(* 상대 PLC 끊김 / 통신 한쪽 고장 *)
_fbRedPeerLost(i_stEntry := TC_EVENTS.PmsSystem.RedPeerLost, i_bActive := i_bRedUse AND i_ePeer = E_RedPeer.Lost, i_nArgs := 0, i_asArg := _asArg);
IF _fbRedLinkFault.q_bRaised <> (i_bRedUse AND (i_ePeer = E_RedPeer.EapLost OR i_ePeer = E_RedPeer.WireLost)) THEN
	IF i_ePeer = E_RedPeer.EapLost THEN
		_asArg[1] := "EAP";
	ELSE
		_asArg[1] := "접점";
	END_IF
END_IF
_fbRedLinkFault(i_stEntry := TC_EVENTS.PmsSystem.RedLinkFault, i_bActive := i_bRedUse AND (i_ePeer = E_RedPeer.EapLost OR i_ePeer = E_RedPeer.WireLost), i_nArgs := 1, i_asArg := _asArg);

(* 동기화 값을 못 받음: EAP는 살아 있는데 동기화 값이 5 s 넘게 안 옴 *)
_tonRedSync(IN := i_bRedUse AND i_bPeerEapOk AND NOT i_bSyncFresh, PT := T#5S);
_fbRedSyncLost(i_stEntry := TC_EVENTS.PmsSystem.RedSyncLost, i_bActive := _tonRedSync.Q, i_nArgs := 0, i_asArg := _asArg);

(* 이중화 설정 오류: 두 PLC 역할이 같거나 Net ID가 RED_SET과 안 맞음 *)
IF _fbRedFailed.q_bRaised <> (i_eRedState = E_RedState.Failed) THEN
	IF i_bRoleConflict THEN
		_asArg[1] := "두 PLC의 역할이 같음";
	ELSE
		_asArg[1] := "이 PLC의 Net ID가 RED_SET과 맞지 않음";
	END_IF
END_IF
_fbRedFailed(i_stEntry := TC_EVENTS.PmsSystem.RedFailed, i_bActive := i_eRedState = E_RedState.Failed, i_nArgs := 1, i_asArg := _asArg);

(* 동기화로 설정을 맞춤 (Active가 바꾼 설정이 이 PLC에 반영됨) *)
IF i_nSyncApplied <> _nRedAppliedLast THEN
	_asArg[1] := TO_WSTRING(i_nSyncApplied - _nRedAppliedLast);
	_nRedAppliedLast := i_nSyncApplied;
	_fbRedSyncApplied.M_SendEvent(1, _asArg);
END_IF
END_ACTION

ACTION A_LogProtection:
// 보호 알람
(* ===== 1) 보호 (알람: 발생·해소 1회씩). 규칙 칸·대상마다. 심각도는 처음 만들 때 조치 기준 ===== *)
FOR _i := 1 TO GVL_PARAM.RULE_COUNT DO
	_m := 0;
	IF iq_aipRule[_i] <> 0 THEN _m := iq_aipRule[_i].ModuleId; END_IF
	FOR _t := 1 TO GVL_PARAM.PROT_TARGET_MAX DO
		// [결함 8 수정 2026-11-03: 대응 칸이 비면 조치가 안 걸리므로 문구·심각도도 조치 없음 (알람만). 원래는 설정 stProt를 그대로 씀:
		//   M_FillProtArgs(..., iq_astRuleCfg[_i].stProt, _asArg) / M_ProtEventBySeverity(iq_astRuleCfg[_i].stProt)]
		_stProtTxt := iq_astRuleCfg[_i].stProt;
		IF iq_aipResp[_i] = 0 THEN
			_stProtTxt.ePcsAction	:= E_PcsAction.None;
			_stProtTxt.eBatAction	:= E_BatAction.None;
			_stProtTxt.eModeAction	:= E_ModeAction.None;
			_stProtTxt.fPPct		:= 100.0;
			_stProtTxt.fQPct		:= 100.0;
		END_IF
		IF _aafbRule[_i, _t].q_bRaised <> iq_aabRule[_i, _t] THEN
			M_FillProtArgs(_m, M_RuleTarget(iq_astRuleCfg[_i].eScope, _t), _stProtTxt, _asArg);
		END_IF
		_aafbRule[_i, _t](i_stEntry := M_ProtEventBySeverity(_stProtTxt), i_bActive := iq_aabRule[_i, _t], i_nArgs := 5, i_asArg := _asArg);
	END_FOR
END_FOR

(* ===== BMS 명령 실패 (알람, 잠그지 않음). 이벤트 항목은 PmsProt.BatLocked를 씀 (문구는 이벤트 클래스에서) ===== *)
FOR _m := 1 TO GVL_PARAM.BMS_COUNT DO
	IF _afbBmsCmdFail[_m].q_bRaised <> (iq_aeBmsFailCmd[_m] <> E_BatCmd.None) THEN
		_asArg[1] := TO_WSTRING(_m);
		_asArg[2] := WCONCAT(F_TxtBatCmd(iq_aeBmsFailCmd[_m]), " 명령 접수 안 됨");
	END_IF
	_afbBmsCmdFail[_m](i_stEntry := TC_EVENTS.PmsProt.BatLocked, i_bActive := iq_aeBmsFailCmd[_m] <> E_BatCmd.None, i_nArgs := 2, i_asArg := _asArg);
END_FOR

(* ===== 가상신호 (알람): 종류가 바뀌면(전압 → 유효전력 등) 해소 후 새 종류로 다시 발생 ===== *)
FOR _g := 1 TO GVL_PARAM.GROUP_COUNT DO
	_nVirtualKind := SEL(i_bTestMode AND iq_astVirtual[_g].bVEna, 0, 1) + SEL(i_bTestMode AND iq_astVirtual[_g].bPEna, 0, 2);
	IF _nVirtualKind <> _anVirtualKind[_g] THEN
		IF _afbVirtual[_g].q_bRaised THEN
			_afbVirtual[_g](i_stEntry := TC_EVENTS.PmsOutput.VirtualOn, i_bActive := FALSE, i_nArgs := 0, i_asArg := _asArg);
		END_IF
		_asArg[1] := TO_WSTRING(_g);
		CASE _nVirtualKind OF
			1:	_asArg[2] := "전압";
			2:	_asArg[2] := "유효전력";
			3:	_asArg[2] := "전압·유효전력";
		END_CASE
		_anVirtualKind[_g] := _nVirtualKind;
	END_IF
	_afbVirtual[_g](i_stEntry := TC_EVENTS.PmsOutput.VirtualOn, i_bActive := _nVirtualKind <> 0, i_nArgs := 2, i_asArg := _asArg);
END_FOR

// 보호가 요청 모드를 Manual로 바꿈 (메시지, 보호가 걸릴 때마다 1회. 걸려 있는 동안 Auto 재요청을 되돌려도 다시 남기지 않음)
FOR _u := 1 TO GVL_PARAM.UNIT_COUNT DO
	IF iq_abModeForced[_u] AND NOT _abModeForcedLogged[_u] THEN
		_asArg[1] := TO_WSTRING(_u);
		_asArg[2] := M_ModuleName(iq_astUnitProt[_u].nModeModule);
		_asArg[3] := TO_WSTRING(iq_astUnitProt[_u].nModeModule);
		_fbModeForced.M_SendEvent(3, _asArg);
		_abModeForcedLogged[_u] := TRUE;
	END_IF
	IF NOT iq_astUnitProt[_u].bModeManualReq THEN
		_abModeForcedLogged[_u] := FALSE;
	END_IF
END_FOR
END_ACTION

ACTION A_LogDeviceFail:
// 명령 실패·장비 쓰기 실패
(* ===== 2) 명령 실패 (알람) ===== *)
FOR _u := 1 TO GVL_PARAM.UNIT_COUNT DO
	IF _afbCmdFail[_u].q_bRaised <> (iq_aeFailCmd[_u] <> E_PcsCmd.None) THEN
		_asArg[1] := TO_WSTRING(_u);
		_asArg[2] := F_TxtPcsCmd(iq_aeFailCmd[_u]);
	END_IF
	_afbCmdFail[_u](i_stEntry := TC_EVENTS.PmsSeq.CmdFail, i_bActive := iq_aeFailCmd[_u] <> E_PcsCmd.None, i_nArgs := 2, i_asArg := _asArg);
END_FOR

(* ===== 2-0) 장비 쓰기 실패 (알람): 드라이버가 상태 bWriteFail로 알림 (FB_DeviceBase.M_MarkWriteResult) ===== *)
FOR _u := 1 TO GVL_PARAM.UNIT_COUNT DO
	IF _afbUnitWriteFail[_u].q_bRaised <> iq_astUnit[_u].bWriteFail THEN
		_asArg[1] := F_TxtNum("유닛 ", _u);
	END_IF
	_afbUnitWriteFail[_u](i_stEntry := TC_EVENTS.PmsSystem.WriteFail, i_bActive := iq_astUnit[_u].bWriteFail, i_nArgs := 1, i_asArg := _asArg);
END_FOR
FOR _m := 1 TO GVL_PARAM.BMS_COUNT DO
	IF _afbBmsWriteFail[_m].q_bRaised <> iq_astBms[_m].bWriteFail THEN
		_asArg[1] := F_TxtNum("BMS ", _m);
	END_IF
	_afbBmsWriteFail[_m](i_stEntry := TC_EVENTS.PmsSystem.WriteFail, i_bActive := iq_astBms[_m].bWriteFail, i_nArgs := 1, i_asArg := _asArg);
END_FOR
END_ACTION

ACTION A_LogSource:
// 지령원 요청·끊김, 코어 상태 요청
(* ===== 3) 지령원: 상태 변경 요청(메시지), 끊김(알람) ===== *)
FOR _i := 1 TO GVL_PARAM.SOURCE_COUNT DO
	IF iq_aipSource[_i] <> 0 AND_THEN iq_astSrcOut[_i].bValid THEN
		_asArg[1] := STRING_TO_WSTRING(iq_aipSource[_i].ModuleName);
		_asArg[2] := TO_WSTRING(iq_aipSource[_i].ModuleId);
		// PCS 요청: 받은 것은 지금 요청과 다를 때만(Reset은 항상), 운전 모드 설정 때문에 무시한 것은 지령 무시로
		IF iq_astSrcOut[_i].stPcsReq.eCmd <> E_PcsCmd.None THEN
			_asArg[3] := F_TxtPcsCmd(iq_astSrcOut[_i].stPcsReq.eCmd);
			IF iq_astSrcOut[_i].stPcsReq.nUnit = 0 THEN
				_asArg[4] := "전체";
			ELSE
				_asArg[4] := F_TxtNum("유닛 ", iq_astSrcOut[_i].stPcsReq.nUnit);
			END_IF
			IF iq_abPcsReqTaken[_i] OR iq_astSrcOut[_i].stPcsReq.eCmd = E_PcsCmd.Reset THEN
				IF iq_astSrcOut[_i].stPcsReq.eCmd <> _aeLastPcsReq[_i] OR iq_astSrcOut[_i].stPcsReq.nUnit <> _anLastPcsUnit[_i]
					OR iq_astSrcOut[_i].stPcsReq.eCmd = E_PcsCmd.Reset THEN
					_fbStateReq.M_SendEvent(4, _asArg);
					_aeLastPcsReq[_i]	:= iq_astSrcOut[_i].stPcsReq.eCmd;
					_anLastPcsUnit[_i]	:= iq_astSrcOut[_i].stPcsReq.nUnit;
				END_IF
			ELSIF i_stSet.bCmdRefused THEN
				_asArg[3] := WCONCAT(_asArg[3], WCONCAT(" ", _asArg[4]));
				_asArg[4] := "이 운전 모드에서 받지 않음 (stStateMode·모드 전환)";
				_fbCmdRefused.M_SendEvent(4, _asArg);
			END_IF
		END_IF
		// 배터리 요청: 받은 것은 항상, 무시한 것은 지령 무시로. Reset은 운전 모드와 관계없이 시퀀서가 보내므로 받은 것으로 기록 (PCS Reset과 같음)
		IF iq_astSrcOut[_i].stBatReq.eCmd <> E_BatCmd.None THEN
			_asArg[3] := F_TxtBatCmd(iq_astSrcOut[_i].stBatReq.eCmd);
			IF iq_astSrcOut[_i].stBatReq.nBatGroup = 0 THEN
				_asArg[4] := "전체";
			ELSE
				_asArg[4] := F_TxtNum("배터리 그룹 ", iq_astSrcOut[_i].stBatReq.nBatGroup);
			END_IF
			IF iq_abBatReqTaken[_i] OR iq_astSrcOut[_i].stBatReq.eCmd = E_BatCmd.Reset THEN
				_fbStateReq.M_SendEvent(4, _asArg);
			ELSIF i_stSet.bCmdRefused THEN
				_asArg[3] := WCONCAT(_asArg[3], WCONCAT(" ", _asArg[4]));
				_asArg[4] := "이 운전 모드에서 받지 않음 (stStateMode)";
				_fbCmdRefused.M_SendEvent(4, _asArg);
			END_IF
		END_IF
	END_IF

	IF iq_astSrcOut[_i].bValid THEN
		_abEverValid[_i] := TRUE;
	END_IF
	// [9번 수정 2026-11-09: 등록 bLostAlarm FALSE면 알람 안 냄 (EMS → 브로커 끊김 알람으로 대신). 원래 조건에 bLostAlarm 없음]
	_bLost := iq_aipSource[_i] <> 0 AND_THEN (iq_astReg[_i].bEnable AND iq_astReg[_i].bLostAlarm AND _abEverValid[_i] AND NOT iq_astSrcOut[_i].bValid);
	IF _afbSrcLost[_i].q_bRaised <> _bLost AND iq_aipSource[_i] <> 0 THEN
		_asArg[1] := STRING_TO_WSTRING(iq_aipSource[_i].ModuleName);
		_asArg[2] := TO_WSTRING(iq_aipSource[_i].ModuleId);
	END_IF
	_afbSrcLost[_i](i_stEntry := TC_EVENTS.PmsOutput.SourceLost, i_bActive := _bLost, i_nArgs := 2, i_asArg := _asArg);
END_FOR
END_ACTION

ACTION A_LogRefused:
// 무시한 지령·기동 조건 대기·지령값 이상·배터리 요청 거부
(* ===== 3-2) 무시한 지령 (메시지): 이상값(지령원별), 방향 반대(유닛별). 새로 생길 때 1회 ===== *)
FOR _i := 1 TO GVL_PARAM.SOURCE_COUNT DO
	IF i_stSet.bCmdRefused AND iq_abBadValue[_i] AND NOT _abLastBad[_i] AND iq_aipSource[_i] <> 0 THEN
		_asArg[1] := STRING_TO_WSTRING(iq_aipSource[_i].ModuleName);
		_asArg[2] := TO_WSTRING(iq_aipSource[_i].ModuleId);
		_asArg[3] := "지령값";
		// [결함 9 수정 2026-11-03: NaN을 비교하지 않고 비트로 봄 (원래 IF iq_afBadValue[_i] <> iq_afBadValue[_i] THEN → FPU 예외)]
		MEMCPY(ADR(_dwBadBits), ADR(iq_afBadValue[_i]), SIZEOF(_dwBadBits));
		IF (_dwBadBits AND 16#7F800000) = 16#7F800000 AND (_dwBadBits AND 16#007FFFFF) <> 0 THEN
			_asArg[4] := "이상값 (숫자 아님)";
		ELSIF (_dwBadBits AND 16#7F800000) = 16#7F800000 OR_ELSE ABS(iq_afBadValue[_i]) >= 1.0E9 THEN
			_asArg[4] := "이상값 (너무 큼)";
		ELSE
			_asArg[4] := WCONCAT("이상값 ", TO_WSTRING(F_RealToDint(iq_afBadValue[_i])));	// [결함 13 수정 2026-11-04: REAL_TO_DINT → F_RealToDint]
		END_IF
		_fbCmdRefused.M_SendEvent(4, _asArg);
	END_IF
	_abLastBad[_i] := iq_abBadValue[_i];
END_FOR
FOR _u := 1 TO GVL_PARAM.UNIT_COUNT DO
	IF i_stSet.bCmdRefused AND iq_aeManualRefuse[_u] <> _aeLastCmdRefuse[_u] AND iq_aeManualRefuse[_u] = E_CmdRefuse.Reversed THEN
		_asArg[1] := M_ModuleName(iq_anManualRefuseModule[_u]);
		_asArg[2] := TO_WSTRING(iq_anManualRefuseModule[_u]);
		_asArg[3] := F_TxtNum("유닛 ", _u);
		_asArg[4] := "방향 반대 (운전 중인 방향과 다름, 앞 값 유지)";
		_fbCmdRefused.M_SendEvent(4, _asArg);
	END_IF
	_aeLastCmdRefuse[_u] := iq_aeManualRefuse[_u];
END_FOR

(* ===== 3-2-1) 기동 조건 대기 (메시지): 대기가 시작되거나 막은 모듈·이유가 바뀔 때 1회 ===== *)
FOR _g := 1 TO GVL_PARAM.GROUP_COUNT DO
	IF iq_abWaitPermit[_g] AND NOT iq_abPermit[_g] THEN
		IF NOT _abPermitLogged[_g] OR iq_anPermitModule[_g] <> _anPermitModule[_g] OR iq_anPermitReason[_g] <> _anPermitReason[_g] THEN
			_asArg[1] := TO_WSTRING(_g);
			_asArg[2] := M_ModuleName(iq_anPermitModule[_g]);
			_asArg[3] := M_ReasonText(iq_anPermitModule[_g], iq_anPermitReason[_g]);
			_asArg[4] := TO_WSTRING(iq_anPermitModule[_g]);
			_fbPermitWait.M_SendEvent(4, _asArg);
			_abPermitLogged[_g]	:= TRUE;
			_anPermitModule[_g]	:= iq_anPermitModule[_g];
			_anPermitReason[_g]	:= iq_anPermitReason[_g];
		END_IF
	ELSE
		_abPermitLogged[_g] := FALSE;
	END_IF
END_FOR

(* ===== 3-2-2) 지령값 이상 (메시지): 디스패처가 NaN·무한대를 0으로 바꾼 유닛, 생길 때 1회 ===== *)
FOR _u := 1 TO GVL_PARAM.UNIT_COUNT DO
	IF iq_abBadSet[_u] AND NOT _abLastBadSet[_u] THEN
		_asArg[1] := TO_WSTRING(_u);
		_fbBadSet.M_SendEvent(1, _asArg);
	END_IF
	_abLastBadSet[_u] := iq_abBadSet[_u];
END_FOR

(* ===== 3-3) 배터리 요청 거부 (메시지): 거부된 요청마다 1회 ===== *)
FOR _b := 1 TO GVL_PARAM.BAT_COUNT DO
	IF i_stSet.bBatRefused AND iq_abBatRefusedNow[_b] THEN
		_asArg[1] := F_TxtNum("배터리 그룹 ", _b);
		IF iq_aeBatRefuse[_b] = E_SeqRefuse.UnitRunning THEN
			_asArg[2] := "배터리 개방";
			_asArg[3] := "버스의 유닛이 운전 중 (정지 후 개방)";
		ELSE
			_asArg[2] := "배터리";
			_asArg[3] := F_TxtRefuse(iq_aeBatRefuse[_b]);
		END_IF
		_fbRefused.M_SendEvent(3, _asArg);
	END_IF
END_FOR
END_ACTION

ACTION A_LogOutput:
// 출력 제한, 자세한 기록
(* ===== 4) 출력 제한: 이유(단계·모듈·이유)가 바뀌고 유지 시간이 지나야 기록 ===== *)
FOR _g := 1 TO GVL_PARAM.GROUP_COUNT DO
	IF NOT M_SameLimitReason(iq_astAutoPDiag[_g], _astCand[_g]) THEN
		_astCand[_g] := iq_astAutoPDiag[_g];
		_atonHold[_g](IN := FALSE);
	END_IF
	_atonHold[_g](IN := NOT M_SameLimitReason(_astCand[_g], _astLogged[_g]), PT := i_stSet.tHold);
	IF _atonHold[_g].Q THEN
		IF M_IsLoggedStage(_astCand[_g].eStage) THEN
			_asArg[1] := TO_WSTRING(_g);
			_asArg[2] := F_TxtStage(_astCand[_g].eStage);
			IF _astCand[_g].eStage = E_DiagStage.UnitLimit THEN
				_asArg[3] := F_TxtLimitBy(_astCand[_g].eUnitBy);
			ELSE
				_asArg[3] := M_ReasonText(_astCand[_g].nModule, _astCand[_g].nReason);
			END_IF
			_asArg[4] := TO_WSTRING(_astCand[_g].nModule);
			_asArg[5] := TO_WSTRING(F_RealToDint(iq_astAutoPDiag[_g].fReq));	// [결함 13 수정 2026-11-04: REAL_TO_DINT → F_RealToDint (NaN·범위 밖 예외 없음)]
			_asArg[6] := TO_WSTRING(F_RealToDint(iq_astAutoPDiag[_g].fOut));
			_fbLimited.M_SendEvent(6, _asArg);
		ELSIF M_IsLoggedStage(_astLogged[_g].eStage) THEN
			_asArg[1] := TO_WSTRING(_g);
			_fbFree.M_SendEvent(1, _asArg);
		END_IF
		_astLogged[_g] := _astCand[_g];
		_atonHold[_g](IN := FALSE);
	END_IF
END_FOR

(* ===== 5) 자세한 기록 (설정으로 켬) ===== *)
FOR _u := 1 TO GVL_PARAM.UNIT_COUNT DO
	IF i_stSet.bUnitLimited AND iq_astUnitDiag[_u].ePBy <> _aeLastLimBy[_u]
		AND iq_astUnitDiag[_u].ePBy <> E_UnitLimitBy.NotRun AND iq_astUnitDiag[_u].ePBy <> E_UnitLimitBy.NotAvail THEN
		_asArg[1] := TO_WSTRING(_u);
		_asArg[2] := F_TxtLimitBy(iq_astUnitDiag[_u].ePBy);
		_asArg[3] := TO_WSTRING(F_RealToDint(iq_astUnitDiag[_u].fPReq));	// [결함 13 수정 2026-11-04: REAL_TO_DINT → F_RealToDint]
		_asArg[4] := TO_WSTRING(F_RealToDint(iq_astUnitDiag[_u].fPOut));
		_fbUnitLim.M_SendEvent(4, _asArg);
	END_IF
	_aeLastLimBy[_u] := iq_astUnitDiag[_u].ePBy;

	IF i_stSet.bReqRefused AND iq_aeRefuse[_u] <> _aeLastRefuse[_u] AND iq_aeRefuse[_u] <> E_SeqRefuse.None THEN
		_asArg[1] := F_TxtNum("유닛 ", _u);
		_asArg[2] := "기동";
		_asArg[3] := F_TxtRefuse(iq_aeRefuse[_u]);
		_fbRefused.M_SendEvent(3, _asArg);
	END_IF
	_aeLastRefuse[_u] := iq_aeRefuse[_u];

	IF i_stSet.bSeqChange AND iq_aeUnitSeq[_u] <> _aeLastSeq[_u] THEN
		_asArg[1] := TO_WSTRING(_u);
		_asArg[2] := F_TxtSeq(_aeLastSeq[_u]);
		_asArg[3] := F_TxtSeq(iq_aeUnitSeq[_u]);
		_fbSeqChange.M_SendEvent(3, _asArg);
	END_IF
	_aeLastSeq[_u] := iq_aeUnitSeq[_u];

	IF i_stSet.bModeChange AND iq_aeOpMode[_u] <> _aeLastMode[_u] THEN
		_asArg[1] := TO_WSTRING(_u);
		_asArg[2] := F_TxtOpMode(_aeLastMode[_u]);
		_asArg[3] := F_TxtOpMode(iq_aeOpMode[_u]);
		_fbModeChange.M_SendEvent(3, _asArg);
	END_IF
	_aeLastMode[_u] := iq_aeOpMode[_u];
END_FOR
END_ACTION

END_FUNCTION_BLOCK

// ---- 10_Core/30_Request/FB_CtrlModeMgr.TcPOU
FUNCTION_BLOCK FB_CtrlModeMgr EXTENDS FB_SourceBase		// 제어 모드 관리자: 등록한 제어 모드(I_ControlMode) 중 하나만 켜고 전환을 맡음. 코어에는 지령원 하나로 보임
// 등록: GVL_SITE.g_aipSource 한 칸 + GVL_PERSIST.g_astSourceReg 같은 칸 (ePowerMode := Auto → Auto 유닛에만 적용). 상태 요청(Run·Stop 등)·제한은 내지 않음
// 요청(i_nModeReq = 모드 칸 번호, 0 = 모드 없음)이 바뀌면: 진입 검사 → 지금 모드 M_Exit → (출력 0 → 지연) → 진입 검사 다시 → 새 모드 M_Enter. 시작한 전환은 끝까지 진행
// 진입 검사에 걸리면 지금 모드를 그대로 둠. 켜진 모드가 스스로 끝내면(bExitReq) 대체 모드(i_stSet.nFallback)로
// 처리한 요청값은 다시 처리하지 않음 (거부·스스로 끝남 뒤 저절로 다시 들어가지 않게). 같은 값을 다시 시도하려면 i_bRetry
// 단위: i_nUnit = 0 → 그룹 하나를 맡음 (그룹 지령 fPSet, 모드는 그룹 값을 봄. 그룹이 2개 이상이면 그룹마다 인스턴스, 등록표 nGroup)
//       i_nUnit = n → 유닛(PCS) n만 맡음 (유닛별 값 astUnit[n], 모드는 FB_UnitView 유닛 값을 봄). PCS마다 관리자 하나 + 모드 인스턴스 한 세트 + 설정 한 세트
//       유닛 단위의 접속점 값은 i_stSet.ePccShare (같은 접속점을 여러 유닛이 쓰면 몫으로 나눔). 접속점이 따로면 유닛마다 제어 그룹을 따로 둠 (GVL_SITE.GROUP_CFG)
// 모드는 FB_ModuleList에 없으므로 설정 점검(M_CheckSet)은 이 FB가 대신 부름
VAR_INPUT
	i_aipMode	: ARRAY[1..GVL_PARAM.CTRL_MODE_COUNT] OF I_ControlMode;	// 등록한 제어 모드 (MAIN 액션 A_PassModuleSet이 GVL_SITE.g_aipCtrlModeN을 매 스캔 넘김). 빈 칸 = 0
	i_stSet		: ST_CtrlModeSet;	// 전환 설정 (A_PassModuleSet이 GVL_PERSIST.g_stModuleSet 칸을 매 스캔 넘김)
	i_nModeReq	: UINT;				// 요청 모드 칸 번호. 0 = 모드 없음 (지령을 내지 않음)
	i_bRetry	: BOOL;				// 같은 요청값을 다시 처리 (쓰면 한 번 처리하고 FALSE로 돌아감)
	i_stTime	: ST_LocalTime;		// 현지 시각 (MAIN 액션 A_PassModuleSet이 매 스캔 넘김). 시간표를 쓰는 모드가 봄
	i_nUnit		: UINT;				// 0 = 그룹 단위. 1~ = 이 유닛(PCS) 단위. 선언에서 정함 (GVL_SITE)
	i_pUnitView	: POINTER TO ARRAY[1..GVL_PARAM.UNIT_COUNT] OF ST_UnitView;	// 유닛 단위일 때: MAIN.fbUnitView.q_astView 주소 (A_PassModuleSet이 매 스캔 넘김). 0 = 연결 안 됨
END_VAR
VAR_OUTPUT
	q_nActive		: UINT;					// 켜진 모드 칸 번호. 0 = 없음 (전환 중에도 0)
	q_sActive		: STRING(31);			// 켜진 모드 이름 (ModuleName)
	q_eStep			: E_CtrlModeStep;		// 관리자 단계
	q_nTarget		: UINT;					// 전환 중 목표 칸 번호 (Leaving일 때만, 0 = 모드 없음으로 가는 중)
	q_eRefuse		: E_CtrlModeRefuse;		// 마지막으로 처리한 요청의 결과 (None = 접수)
	q_nRefuseReason	: UINT;					// NotReady일 때 그 모드의 이유 코드 (M_ModeReasonText)
	q_nExitSlot		: UINT;					// 마지막으로 스스로 끝낸 모드 칸 번호
	q_nExitReason	: UINT;					// 그 이유 코드 (M_ModeReasonText)
	q_bChanged		: BOOL;					// 켜진 모드가 바뀐 스캔 (1스캔, 기록용)
	q_bRefusedNow	: BOOL;					// 이번 스캔에 요청을 거부함 (1스캔, 기록용). 칸 q_nRefuseSlot, 결과 q_eRefuse·q_nRefuseReason [7번 수정 2026-11-09: 추가]
	q_nRefuseSlot	: UINT;					// 마지막으로 거부한 요청 칸 번호
	q_bExitedNow	: BOOL;					// 이번 스캔에 켜진 모드가 스스로 끝남 (1스캔, 기록용). 칸 q_nExitSlot, 이유 q_nExitReason [7번 수정 2026-11-09: 추가]
	q_fPccP			: REAL;					// kW, 모드가 본 접속점 P (공급 +). 유닛 단위면 ePccShare를 적용한 값
END_VAR
VAR
	_nHandledReq	: UINT;				// 처리를 끝낸 요청값 (요청이 이것과 다를 때만 새로 처리)
	_nActive		: UINT;				// 켜진 모드 칸 번호
	_nTarget		: UINT;				// 진행 중인 전환의 목표 (끝날 때까지 고정)
	_bLeaveP		: BOOL;				// 전환 중 P를 0으로 냄 (이전 모드가 P를 내던 경우만)
	_bLeaveQ		: BOOL;				// 전환 중 Q를 0으로 냄
	_bPrevP			: BOOL;				// 켜진 모드가 지난 스캔에 P를 냄
	_bPrevQ			: BOOL;
	_tonZero		: TON;
	_stModeOut		: ST_CtrlModeOut;	// 켜진 모드의 이번 스캔 결과
	_stModeView		: ST_CtrlModeView;	// 모드에 넘기는 값 (이번 스캔)
	(* [16번 수정 2026-11-09: 추가] 유닛별 값을 내는 모드(bUnitOut)의 전환 중 0 *)
	_bPrevUnitOut	: BOOL;				// 켜진 모드가 지난 스캔에 유닛별 값을 냄
	_abPrevUnitP	: ARRAY[1..GVL_PARAM.UNIT_COUNT] OF BOOL;
	_abPrevUnitQ	: ARRAY[1..GVL_PARAM.UNIT_COUNT] OF BOOL;
	_bLeaveUnit		: BOOL;				// 전환 중 유닛 칸으로 0을 냄 (이전 모드가 유닛별 값을 내던 경우)
	_abLeaveUnitP	: ARRAY[1..GVL_PARAM.UNIT_COUNT] OF BOOL;
	_abLeaveUnitQ	: ARRAY[1..GVL_PARAM.UNIT_COUNT] OF BOOL;
END_VAR

METHOD M_UpdateOutput : BOOL
VAR
	stNoMode	: ST_CtrlModeOut;
	stOld		: ST_SourceOutput;	// 지난 스캔 낸 값 (새 지령 판단)
	bNew		: BOOL;
	stNoReq		: ST_UnitReq;
	k			: UINT;
	nCode		: UINT;
	nFallback	: UINT;
	bOk			: BOOL;
END_VAR
q_bChanged	:= FALSE;
q_bRefusedNow	:= FALSE;
q_bExitedNow	:= FALSE;
IF i_nUnit = 0 THEN
	_stModeView.stGroup	:= _stView;		// FB_SourceBase가 이번 스캔 채운 대상 그룹 값
ELSE
	_stModeView.stGroup	:= M_UnitView();	// 이 유닛 값 (접속점은 ePccShare 몫)
END_IF
_stModeView.stTime	:= i_stTime;
q_fPccP := _stModeView.stGroup.stPcc.stMeas.stP.fValue;

// 0) 켜진 모드가 등록에서 빠졌으면 (온라인 변경) 모드 없음으로
IF q_eStep = E_CtrlModeStep.Active AND NOT M_Valid(i_nSlot := _nActive) THEN
	_nActive	:= 0;
	q_eStep		:= E_CtrlModeStep.Idle;
	q_bChanged	:= TRUE;
END_IF

// 1) 새 요청 (전환 중이면 끝난 뒤 처리)
IF q_eStep <> E_CtrlModeStep.Leaving AND (i_nModeReq <> _nHandledReq OR i_bRetry) THEN
	_nHandledReq	:= i_nModeReq;
	q_eRefuse		:= E_CtrlModeRefuse.None;
	q_nRefuseReason	:= 0;
	IF i_nModeReq <> _nActive THEN
		IF i_nModeReq <> 0 AND NOT M_Valid(i_nSlot := i_nModeReq) THEN
			q_eRefuse := E_CtrlModeRefuse.BadSlot;
			q_nRefuseSlot	:= i_nModeReq;
			q_bRefusedNow	:= TRUE;
		ELSE
			nCode := 0;
			IF i_nModeReq <> 0 THEN
				nCode := i_aipMode[i_nModeReq].M_CheckEnter(i_stView := _stModeView);
			END_IF
			IF nCode = 0 THEN
				M_StartSwitch(i_nTarget := i_nModeReq);
			ELSE
				q_eRefuse		:= E_CtrlModeRefuse.NotReady;	// 지금 모드는 그대로
				q_nRefuseReason	:= nCode;
				q_nRefuseSlot	:= i_nModeReq;
				q_bRefusedNow	:= TRUE;
			END_IF
		END_IF
	END_IF
	i_bRetry := FALSE;		// 처리한 뒤에만 지움 (전환 중에 온 재시도는 끝난 뒤 처리)
END_IF

// 2) 전환 중: 0으로 둔 시간이 지나면 진입 검사를 다시 하고 새 모드로 (지연 동안 조건이 바뀌었을 수 있음)
_tonZero(IN := q_eStep = E_CtrlModeStep.Leaving, PT := i_stSet.tZeroDelay);
IF q_eStep = E_CtrlModeStep.Leaving AND _tonZero.Q THEN
	bOk := TRUE;
	IF _nTarget <> 0 THEN
		IF M_Valid(i_nSlot := _nTarget) THEN
			nCode := i_aipMode[_nTarget].M_CheckEnter(i_stView := _stModeView);
			IF nCode <> 0 THEN
				bOk				:= FALSE;
				q_eRefuse		:= E_CtrlModeRefuse.NotReady;
				q_nRefuseReason	:= nCode;
			END_IF
		ELSE
			bOk				:= FALSE;
			q_eRefuse		:= E_CtrlModeRefuse.BadSlot;
			q_nRefuseReason	:= 0;
		END_IF
		IF NOT bOk THEN
			q_nRefuseSlot	:= _nTarget;
			q_bRefusedNow	:= TRUE;
		END_IF
	END_IF
	IF bOk THEN
		M_EnterMode(i_nSlot := _nTarget);
	ELSE
		M_EnterMode(i_nSlot := 0);
	END_IF
END_IF

// 3) 켜진 모드 계산. 스스로 끝내면 대체 모드로
IF q_eStep = E_CtrlModeStep.Active THEN
	_bPrevP		:= _stModeOut.bPSetActive;		// 지난 스캔에 내던 쪽 (끝내는 스캔에 지령을 비워도 0으로 둘 수 있게)
	_bPrevQ		:= _stModeOut.bQSetActive;
	_bPrevUnitOut	:= _stModeOut.bUnitOut;
	FOR k := 1 TO GVL_PARAM.UNIT_COUNT DO
		_abPrevUnitP[k]	:= _stModeOut.bUnitOut AND _stModeOut.astUnit[k].bPSetActive;
		_abPrevUnitQ[k]	:= _stModeOut.bUnitOut AND _stModeOut.astUnit[k].bQSetActive;
	END_FOR
	_stModeOut	:= i_aipMode[_nActive].M_Calc(i_stView := _stModeView);
	IF _stModeOut.bExitReq THEN
		q_nExitSlot		:= _nActive;
		q_nExitReason	:= _stModeOut.nReason;
		q_bExitedNow	:= TRUE;
		nFallback		:= 0;
		IF i_stSet.nFallback <> _nActive AND M_Valid(i_nSlot := i_stSet.nFallback) THEN
			IF i_aipMode[i_stSet.nFallback].M_CheckEnter(i_stView := _stModeView) = 0 THEN
				nFallback := i_stSet.nFallback;
			END_IF
		END_IF
		M_StartSwitch(i_nTarget := nFallback);
		// 대체 모드로 바로 들어갔으면 이번 스캔 값을 냄 (그 모드의 bExitReq는 다음 스캔에 봄)
		IF q_eStep = E_CtrlModeStep.Active THEN
			_stModeOut := i_aipMode[_nActive].M_Calc(i_stView := _stModeView);
		END_IF
	END_IF
ELSIF q_eStep = E_CtrlModeStep.Idle THEN
	_stModeOut	:= stNoMode;
	_bPrevP		:= FALSE;
	_bPrevQ		:= FALSE;
	_bPrevUnitOut	:= FALSE;
	FOR k := 1 TO GVL_PARAM.UNIT_COUNT DO
		_abPrevUnitP[k]	:= FALSE;
		_abPrevUnitQ[k]	:= FALSE;
	END_FOR
END_IF

// 4) 출력: P·Q 지령만 (제한·상태 요청은 내지 않음). 그룹 단위 = 그룹 지령, 유닛 단위 = 그 유닛 칸만
//    [16번 수정 2026-11-09: 모드가 유닛별 값을 내면(bUnitOut, 스탠다드 스케줄) 접속점 그룹 단위에서도 유닛 칸으로 냄 (접속점 그룹 지령은 비움).
//     유닛 단위면 맡은 유닛 칸만. 원래는 모드의 접속점 그룹 값(fPSet·fQSet)만 냄]
// 지난 스캔 값 (FB_SourceBase가 끊김·사용 안 함으로 비웠으면 빈 값과 비교 → 다시 켜질 때 새 지령)
stOld := _stOut;
// 모두 비우고 맡은 칸만 씀 (i_nUnit을 온라인으로 바꿔도 이전 칸이 남지 않게). 범위 밖이면 아무것도 안 냄 (설정 점검 오류)
_stOut.bPSetActive	:= FALSE;
_stOut.fPSet		:= 0.0;
_stOut.bQSetActive	:= FALSE;
_stOut.fQSet		:= 0.0;
FOR k := 1 TO GVL_PARAM.UNIT_COUNT DO
	_stOut.astUnit[k] := stNoReq;
END_FOR
CASE q_eStep OF
	E_CtrlModeStep.Active:
		IF _stModeOut.bUnitOut THEN
			FOR k := 1 TO GVL_PARAM.UNIT_COUNT DO
				IF i_nUnit = 0 OR i_nUnit = k THEN
					_stOut.astUnit[k] := _stModeOut.astUnit[k];
				END_IF
			END_FOR
		ELSIF i_nUnit = 0 THEN
			_stOut.bPSetActive	:= _stModeOut.bPSetActive;
			_stOut.fPSet		:= _stModeOut.fPSet;
			_stOut.bQSetActive	:= _stModeOut.bQSetActive;
			_stOut.fQSet		:= _stModeOut.fQSet;
		ELSIF i_nUnit <= GVL_PARAM.UNIT_COUNT THEN
			_stOut.astUnit[i_nUnit].bPSetActive	:= _stModeOut.bPSetActive;
			_stOut.astUnit[i_nUnit].fPSet		:= _stModeOut.fPSet;
			_stOut.astUnit[i_nUnit].bQSetActive	:= _stModeOut.bQSetActive;
			_stOut.astUnit[i_nUnit].fQSet		:= _stModeOut.fQSet;
		END_IF
	E_CtrlModeStep.Leaving:
		// 이전 모드가 내던 쪽만 0을 냄 (비우면 그 사이 등급이 낮은 지령원 값이 들어옴)
		IF _bLeaveUnit THEN
			FOR k := 1 TO GVL_PARAM.UNIT_COUNT DO
				IF i_nUnit = 0 OR i_nUnit = k THEN
					_stOut.astUnit[k].bPSetActive	:= _abLeaveUnitP[k];
					_stOut.astUnit[k].bQSetActive	:= _abLeaveUnitQ[k];
				END_IF
			END_FOR
		ELSIF i_nUnit = 0 THEN
			_stOut.bPSetActive	:= _bLeaveP;
			_stOut.bQSetActive	:= _bLeaveQ;
		ELSIF i_nUnit <= GVL_PARAM.UNIT_COUNT THEN
			_stOut.astUnit[i_nUnit].bPSetActive	:= _bLeaveP;
			_stOut.astUnit[i_nUnit].bQSetActive	:= _bLeaveQ;
		END_IF
END_CASE
// [결함 13 수정 2026-11-04: 값 비교를 비트로 (모드 출력이 NaN이어도 여기서 멈추지 않고, 고르기(F_CmdOk)에서 이상값으로 거름)]
bNew := _stOut.bPSetActive <> stOld.bPSetActive OR F_RealChanged(_stOut.fPSet, stOld.fPSet)
	OR _stOut.bQSetActive <> stOld.bQSetActive OR F_RealChanged(_stOut.fQSet, stOld.fQSet);
FOR k := 1 TO GVL_PARAM.UNIT_COUNT DO
	bNew := bNew OR _stOut.astUnit[k].bPSetActive <> stOld.astUnit[k].bPSetActive OR F_RealChanged(_stOut.astUnit[k].fPSet, stOld.astUnit[k].fPSet)
		OR _stOut.astUnit[k].bQSetActive <> stOld.astUnit[k].bQSetActive OR F_RealChanged(_stOut.astUnit[k].fQSet, stOld.astUnit[k].fQSet);
END_FOR
_stOut.bNewSet := bNew;

// 5) 진단
q_nActive := _nActive;
q_sActive := '';
IF q_eStep = E_CtrlModeStep.Active THEN
	q_sActive := i_aipMode[_nActive].ModuleName;
END_IF
q_nTarget := 0;
IF q_eStep = E_CtrlModeStep.Leaving THEN
	q_nTarget := _nTarget;
END_IF

M_UpdateOutput := TRUE;		// 관리자는 늘 살아 있음 (만료 없음). 모드가 없으면 지령 없음
END_METHOD

METHOD PRIVATE M_UnitView : ST_GroupView		// 유닛 단위: 이 유닛 값 (FB_UnitView)에 접속점 몫을 적용. 연결 안 됐으면 빈 값 (가용 유닛 0 → 모드 진입 안 됨)
VAR
	stUv		: ST_UnitView;
	stNone		: ST_GroupView;
	fShare		: REAL;
	fLoad		: REAL;
END_VAR
M_UnitView := stNone;
IF i_nUnit < 1 OR i_nUnit > GVL_PARAM.UNIT_COUNT OR i_pUnitView = 0 THEN
	RETURN;		// 설정 점검(M_CheckSet)이 오류로 올림
END_IF
stUv		:= i_pUnitView^[i_nUnit];
M_UnitView	:= stUv.stView;
IF i_stSet.ePccShare = E_PccShare.Actual THEN
	RETURN;		// 접속점 실측 그대로
END_IF
IF i_stSet.ePccShare = E_PccShare.Fixed THEN
	fShare := LIMIT(0.0, i_stSet.fPccRatio, 1.0);
ELSE
	fShare := stUv.fRatingShare;
END_IF
// 모드는 부하를 '출력 - 접속점 P'로 셈. 이 유닛 몫 부하 = 몫 × (그룹 출력 - 접속점 P)가 되도록 접속점 P = 유닛 출력 - 몫 부하
IF stUv.stView.stPcc.stMeas.stP.bValid THEN
	fLoad := stUv.fGroupPOut - stUv.stView.stPcc.stMeas.stP.fValue;
	M_UnitView.stPcc.stMeas.stP.fValue := stUv.stView.fPOut - fShare * fLoad;
END_IF
IF stUv.stView.stPcc.stMeas.stQ.bValid THEN
	fLoad := stUv.fGroupQOut - stUv.stView.stPcc.stMeas.stQ.fValue;
	M_UnitView.stPcc.stMeas.stQ.fValue := stUv.stView.fQOut - fShare * fLoad;
END_IF
END_METHOD

METHOD PRIVATE M_StartSwitch		// 지금 모드를 끝내고 목표로 전환 시작 (0으로 둘 게 있으면 Leaving, 없으면 바로 진입)
VAR_INPUT
	i_nTarget	: UINT;		// 목표 칸 번호. 0 = 모드 없음. 0이 아니면 부르는 쪽이 진입 검사를 마침
END_VAR
VAR
	bWasActive	: BOOL;
	bLeaveAnyUnit	: BOOL;		// 유닛 칸 중 0으로 둘 것이 있음
	k			: UINT;
END_VAR
bWasActive := q_eStep = E_CtrlModeStep.Active;
bLeaveAnyUnit := FALSE;
IF bWasActive THEN
	i_aipMode[_nActive].M_Exit();
	_bLeaveP	:= _stModeOut.bPSetActive OR _bPrevP;		// 이전 모드가 이번·지난 스캔에 내던 쪽
	_bLeaveQ	:= _stModeOut.bQSetActive OR _bPrevQ;
	// [16번 수정 2026-11-09: 유닛별 값을 내던 모드면 유닛 칸마다 같은 방식으로]
	_bLeaveUnit	:= _stModeOut.bUnitOut OR _bPrevUnitOut;
	FOR k := 1 TO GVL_PARAM.UNIT_COUNT DO
		_abLeaveUnitP[k]	:= (_stModeOut.bUnitOut AND _stModeOut.astUnit[k].bPSetActive) OR _abPrevUnitP[k];
		_abLeaveUnitQ[k]	:= (_stModeOut.bUnitOut AND _stModeOut.astUnit[k].bQSetActive) OR _abPrevUnitQ[k];
		bLeaveAnyUnit		:= bLeaveAnyUnit OR _abLeaveUnitP[k] OR _abLeaveUnitQ[k];
	END_FOR
	_nActive	:= 0;
	q_bChanged	:= TRUE;
END_IF
_nTarget := i_nTarget;
IF bWasActive AND i_stSet.bZeroOnSwitch AND (_bLeaveP OR _bLeaveQ OR (_bLeaveUnit AND bLeaveAnyUnit)) THEN
	_tonZero(IN := FALSE);		// 지연을 처음부터 셈
	q_eStep := E_CtrlModeStep.Leaving;
ELSE
	M_EnterMode(i_nSlot := i_nTarget);
END_IF
END_METHOD

METHOD PRIVATE M_EnterMode		// 모드 진입 (0 = 모드 없음으로)
VAR_INPUT
	i_nSlot		: UINT;		// 0이 아니면 등록된 칸이어야 함 (부르는 쪽이 확인)
END_VAR
_nTarget := 0;
IF i_nSlot = 0 THEN
	_nActive	:= 0;
	q_eStep		:= E_CtrlModeStep.Idle;
ELSE
	i_aipMode[i_nSlot].M_Enter(i_stView := _stModeView);
	_nActive	:= i_nSlot;
	q_eStep		:= E_CtrlModeStep.Active;
	q_bChanged	:= TRUE;
END_IF
END_METHOD

METHOD PRIVATE M_Valid : BOOL		// 칸 번호가 범위 안이고 모드가 등록됨
VAR_INPUT
	i_nSlot		: UINT;
END_VAR
// AND는 단락 평가가 아니므로 범위를 먼저 따로 봄 (배열 범위 밖 접근 방지)
M_Valid := FALSE;
IF i_nSlot >= 1 AND i_nSlot <= GVL_PARAM.CTRL_MODE_COUNT THEN
	M_Valid := i_aipMode[i_nSlot] <> 0;
END_IF
END_METHOD

METHOD M_CheckSet : WSTRING(63)		// 대체 모드 칸 번호 + 등록한 모드마다 M_CheckSet (첫 오류 문구)
VAR
	i			: UINT;
	sErr		: WSTRING(63);
END_VAR
M_CheckSet := "";
IF i_nUnit > GVL_PARAM.UNIT_COUNT THEN
	M_CheckSet := "제어 모드: i_nUnit이 유닛 수(UNIT_COUNT)보다 큼";
	RETURN;
END_IF
IF i_nUnit <> 0 AND i_pUnitView = 0 THEN
	M_CheckSet := "제어 모드: 유닛 단위인데 유닛 값(i_pUnitView) 연결 안 됨";
	RETURN;
END_IF
IF NOT F_RealOk(i_stSet.fPccRatio) THEN	// [결함 13 수정 2026-11-04]
	M_CheckSet := "제어 모드: 접속점 몫 fPccRatio 숫자 아님";
	RETURN;
END_IF
IF i_stSet.ePccShare = E_PccShare.Fixed AND NOT (i_stSet.fPccRatio >= 0.0 AND i_stSet.fPccRatio <= 1.0) THEN
	M_CheckSet := "제어 모드: 접속점 몫 fPccRatio는 0~1";
	RETURN;
END_IF
IF i_stSet.nFallback <> 0 AND NOT M_Valid(i_nSlot := i_stSet.nFallback) THEN
	M_CheckSet := "제어 모드: 대체 모드 nFallback 칸이 비었거나 범위 밖";
	RETURN;
END_IF
FOR i := 1 TO GVL_PARAM.CTRL_MODE_COUNT DO
	IF i_aipMode[i] <> 0 THEN
		sErr := i_aipMode[i].M_CheckSet();
		IF sErr <> "" THEN
			M_CheckSet := sErr;
			RETURN;
		END_IF
	END_IF
END_FOR
END_METHOD

METHOD M_SlotName : WSTRING(63)		// 모드 칸 번호 → 이름 (0 = 없음). 로그용 [7번 수정 2026-11-09: 추가]
VAR_INPUT
	i_nSlot		: UINT;
END_VAR
IF i_nSlot = 0 THEN
	M_SlotName := "없음";
ELSIF M_Valid(i_nSlot := i_nSlot) THEN
	M_SlotName := STRING_TO_WSTRING(i_aipMode[i_nSlot].ModuleName);
ELSE
	M_SlotName := WCONCAT("칸 ", TO_WSTRING(i_nSlot));
END_IF
END_METHOD

METHOD M_RefuseText : WSTRING(63)		// 마지막 거부 이유 문구 (q_eRefuse·q_nRefuseSlot·q_nRefuseReason). 로그용 [7번 수정 2026-11-09: 추가]
CASE q_eRefuse OF
	E_CtrlModeRefuse.BadSlot:
		M_RefuseText := "모드 칸이 비었거나 범위 밖";
	E_CtrlModeRefuse.NotReady:
		M_RefuseText := M_ModeReasonText(i_nSlot := q_nRefuseSlot, i_nReason := q_nRefuseReason);
ELSE
	M_RefuseText := "";
END_CASE
END_METHOD

METHOD M_ModeReasonText : WSTRING(63)		// 모드 칸의 이유 코드 → 문구 (q_nRefuseReason·q_nExitReason을 HMI·로그에 보일 때)
VAR_INPUT
	i_nSlot		: UINT;
	i_nReason	: UINT;
END_VAR
IF M_Valid(i_nSlot := i_nSlot) THEN
	M_ModeReasonText := i_aipMode[i_nSlot].M_ReasonText(i_nReason := i_nReason);
ELSE
	M_ModeReasonText := WCONCAT("이유 ", TO_WSTRING(i_nReason));
END_IF
END_METHOD

END_FUNCTION_BLOCK

// ---- 10_Core/03_Base/FB_SourceBase.TcPOU
FUNCTION_BLOCK ABSTRACT FB_SourceBase EXTENDS FB_ModuleBase IMPLEMENTS I_CommandSource
VAR
	_stOut			: ST_SourceOutput;
	_stView			: ST_GroupView;		// 이번 스캔 대상 그룹 값 (파생 FB의 M_UpdateOutput에서 읽음)
	_tonExpire		: TON;
	_bEverAlive		: BOOL;
END_VAR

PROPERTY Output : ST_SourceOutput
GET
Output := _stOut;
END_GET
END_PROPERTY

METHOD M_Cycle
VAR_INPUT
	i_stReg		: ST_SourceReg;
	i_stView	: ST_GroupView;
END_VAR
VAR
	bFresh		: BOOL;
	u			: UINT;
END_VAR
_stView := i_stView;

// 1) 파생 FB가 _stOut을 채운다. 값이 새로 들어왔으면 TRUE
//    상태 요청은 1스캔만: 파생 FB가 새 요청이 있을 때만 다시 채움
_stOut.stPcsReq.eCmd := E_PcsCmd.None;
_stOut.stBatReq.eCmd := E_BatCmd.None;
_stOut.bNewSet := FALSE;		// 새 지령도 1스캔만: 파생 FB가 새 값이 들어왔을 때 TRUE로
bFresh := M_UpdateOutput();
IF bFresh THEN
	_bEverAlive := TRUE;
END_IF
_tonExpire(IN := NOT bFresh, PT := i_stReg.tExpire);

// 2) 공통 처리
IF NOT i_stReg.bEnable OR NOT _bEverAlive THEN
	M_ClearAll();
ELSIF _tonExpire.Q THEN
	// 끊김: 지령·상태 요청은 무효 (그룹·유닛별 모두), 제한(P·Q)은 마지막 값 유지
	_stOut.bPSetActive	:= FALSE;
	_stOut.bQSetActive	:= FALSE;
	_stOut.stPcsReq.eCmd	:= E_PcsCmd.None;
	_stOut.stBatReq.eCmd	:= E_BatCmd.None;
	_stOut.bNewSet		:= FALSE;
	FOR u := 1 TO GVL_PARAM.UNIT_COUNT DO
		_stOut.astUnit[u].bPSetActive := FALSE;
		_stOut.astUnit[u].bQSetActive := FALSE;
	END_FOR
	_stOut.bValid		:= _stOut.bPLimActive OR _stOut.bQLimActive;	// 유지할 제한(P·Q)이 있을 때만 유효
ELSE
	_stOut.bValid := TRUE;
END_IF
END_METHOD

METHOD ABSTRACT M_UpdateOutput : BOOL		// 파생 FB: _stOut을 채우고, 새 값이 들어왔으면 TRUE
END_METHOD

METHOD PROTECTED M_ClearAll
VAR
	stNone		: ST_SourceOutput;
END_VAR
_stOut := stNone;
END_METHOD

METHOD M_ReasonText : WSTRING(63)	// 지령원이 낸 P 제한의 이유 문구 (지령원 제한은 이유 코드를 쓰지 않음)
VAR_INPUT
	i_nReason	: UINT;
END_VAR
M_ReasonText := "지령원 제한";
END_METHOD

END_FUNCTION_BLOCK

// ---- 10_Core/02_Util/F_RealChanged.TcPOU
FUNCTION F_RealChanged : BOOL		// 두 REAL의 비트가 다른가 (새 지령 판단용). NaN이 들어와도 비교 예외 없음 [결함 13 수정 2026-11-04: 추가]
VAR_INPUT
	i_fA		: REAL;
	i_fB		: REAL;
END_VAR
VAR
	dwA			: DWORD;
	dwB			: DWORD;
END_VAR

MEMCPY(ADR(dwA), ADR(i_fA), SIZEOF(dwA));
MEMCPY(ADR(dwB), ADR(i_fB), SIZEOF(dwB));
F_RealChanged := dwA <> dwB;

END_FUNCTION

// ---- 10_Core/70_Diag/F_TxtPcsAction.TcPOU
FUNCTION F_TxtPcsAction : WSTRING(31)		// PCS 조치 문구
VAR_INPUT
	i_e		: E_PcsAction;
END_VAR

CASE i_e OF
	E_PcsAction.None:	F_TxtPcsAction := "알람만";
	E_PcsAction.Standby:	F_TxtPcsAction := "대기";
	E_PcsAction.Stop:	F_TxtPcsAction := "정지";
	E_PcsAction.EStop:	F_TxtPcsAction := "비상정지";
ELSE
	F_TxtPcsAction := "?";
END_CASE

END_FUNCTION

// ---- 10_Core/70_Diag/F_TxtBatAction.TcPOU
FUNCTION F_TxtBatAction : WSTRING(31)		// 배터리 조치 문구
VAR_INPUT
	i_e		: E_BatAction;
END_VAR

CASE i_e OF
	E_BatAction.None:	F_TxtBatAction := "조치 없음";
	E_BatAction.Stop:	F_TxtBatAction := "개방";
	E_BatAction.EStop:	F_TxtBatAction := "비상정지";
ELSE
	F_TxtBatAction := "?";
END_CASE

END_FUNCTION

// ---- 10_Core/70_Diag/F_TxtCoreReason.TcPOU
FUNCTION F_TxtCoreReason : WSTRING(63)		// 코어 제한 이유 문구 (모듈 ID 0)
VAR_INPUT
	i_nReason	: UINT;
END_VAR

IF i_nReason = GVL_REASON.RSN_RATING THEN
	F_TxtCoreReason := "가용 유닛 정격";
ELSIF i_nReason = GVL_REASON.RSN_BAT THEN
	F_TxtCoreReason := "배터리 충·방전 한도";
ELSIF i_nReason = GVL_REASON.RSN_RATING_Q THEN
	F_TxtCoreReason := "가용 유닛 Q 정격";
ELSIF i_nReason = GVL_REASON.RSN_DERATE THEN
	F_TxtCoreReason := "보호 Derate";
ELSE
	F_TxtCoreReason := WCONCAT("코어 이유 ", TO_WSTRING(i_nReason));
END_IF

END_FUNCTION

// ---- 10_Core/70_Diag/F_TxtNum.TcPOU
FUNCTION F_TxtNum : WSTRING(63)		// 앞말 + 번호 (예: "유닛 2")
VAR_INPUT
	i_sPrefix	: WSTRING(47);			// 설정 오류 문구처럼 긴 앞말도 받음
	i_nNum		: UINT;
END_VAR

F_TxtNum := WCONCAT(i_sPrefix, TO_WSTRING(i_nNum));

END_FUNCTION

// ---- 10_Core/70_Diag/F_TxtBatCmd.TcPOU
FUNCTION F_TxtBatCmd : WSTRING(31)
VAR_INPUT
	i_e		: E_BatCmd;
END_VAR

CASE i_e OF
	E_BatCmd.None:		F_TxtBatCmd := "없음";
	E_BatCmd.Close:		F_TxtBatCmd := "배터리 투입";
	E_BatCmd.Open:		F_TxtBatCmd := "배터리 개방";
	E_BatCmd.EStop:		F_TxtBatCmd := "배터리 비상정지";
	E_BatCmd.Reset:		F_TxtBatCmd := "배터리 Reset";
ELSE
	F_TxtBatCmd := "?";
END_CASE

END_FUNCTION

// ---- 10_Core/70_Diag/F_TxtPcsCmd.TcPOU
FUNCTION F_TxtPcsCmd : WSTRING(31)
VAR_INPUT
	i_e		: E_PcsCmd;
END_VAR

CASE i_e OF
	E_PcsCmd.None:		F_TxtPcsCmd := "없음";
	E_PcsCmd.Run:		F_TxtPcsCmd := "Run";
	E_PcsCmd.Standby:	F_TxtPcsCmd := "Standby";
	E_PcsCmd.Stop:		F_TxtPcsCmd := "Stop";
	E_PcsCmd.Reset:		F_TxtPcsCmd := "Reset";
	E_PcsCmd.EStop:		F_TxtPcsCmd := "EStop";
ELSE
	F_TxtPcsCmd := "?";
END_CASE

END_FUNCTION

// ---- 10_Core/02_Util/F_RealToDint.TcPOU
FUNCTION F_RealToDint : DINT		// REAL → DINT, NaN·무한대는 0, 범위 밖은 끝값으로 (REAL_TO_DINT는 NaN·범위 밖이면 FPU 예외) [결함 13 수정 2026-11-04: 추가]
VAR_INPUT
	i_fValue	: REAL;
END_VAR

IF NOT F_RealOk(i_fValue) THEN
	F_RealToDint := 0;
ELSIF i_fValue >= 2147483520.0 THEN		// REAL로 나타낼 수 있는 DINT 최댓값 근처
	F_RealToDint := 2147483520;
ELSIF i_fValue <= -2147483520.0 THEN
	F_RealToDint := -2147483520;
ELSE
	F_RealToDint := REAL_TO_DINT(i_fValue);
END_IF

END_FUNCTION

// ---- 10_Core/70_Diag/F_TxtRefuse.TcPOU
FUNCTION F_TxtRefuse : WSTRING(31)		// 거부 이유 문구
VAR_INPUT
	i_e		: E_SeqRefuse;
END_VAR

CASE i_e OF
	E_SeqRefuse.None:	F_TxtRefuse := "없음";
	E_SeqRefuse.NotAvail:	F_TxtRefuse := "가용 아님";
	E_SeqRefuse.NoBattery:	F_TxtRefuse := "배터리 미투입";
	E_SeqRefuse.NoPermit:	F_TxtRefuse := "기동 조건 미충족";
	E_SeqRefuse.CommLost:	F_TxtRefuse := "통신 없음";
	E_SeqRefuse.UnitRunning:	F_TxtRefuse := "유닛 운전 중";
	E_SeqRefuse.StopInProgress:	F_TxtRefuse := "정지 진행 중";
	E_SeqRefuse.ConfigError:	F_TxtRefuse := "설정 오류";
	E_SeqRefuse.WriteDisabled:	F_TxtRefuse := "장비 쓰기 불가";
ELSE
	F_TxtRefuse := "?";
END_CASE

END_FUNCTION

// ---- 10_Core/70_Diag/F_TxtStage.TcPOU
FUNCTION F_TxtStage : WSTRING(31)		// 진단 단계 문구
VAR_INPUT
	i_e		: E_DiagStage;
END_VAR

CASE i_e OF
	E_DiagStage.None:	F_TxtStage := "없음";
	E_DiagStage.NoRequest:	F_TxtStage := "요청 없음";
	E_DiagStage.NotRunning:	F_TxtStage := "운전 아님";
	E_DiagStage.Ramp:	F_TxtStage := "램프";
	E_DiagStage.PccLimit:	F_TxtStage := "접속점 제한";
	E_DiagStage.DeviceLimit:	F_TxtStage := "설비 제한";
	E_DiagStage.UnitLimit:	F_TxtStage := "유닛 한도·분배";
	E_DiagStage.NoUnit:	F_TxtStage := "이 모드 유닛 없음";
ELSE
	F_TxtStage := "?";
END_CASE

END_FUNCTION

// ---- 10_Core/70_Diag/F_TxtLimitBy.TcPOU
FUNCTION F_TxtLimitBy : WSTRING(31)		// 유닛 축소 이유 문구
VAR_INPUT
	i_e		: E_UnitLimitBy;
END_VAR

CASE i_e OF
	E_UnitLimitBy.None:	F_TxtLimitBy := "없음";
	E_UnitLimitBy.NotAvail:	F_TxtLimitBy := "가용 아님";
	E_UnitLimitBy.NotRun:	F_TxtLimitBy := "활성 아님·정지 중";
	E_UnitLimitBy.Rating:	F_TxtLimitBy := "정격";
	E_UnitLimitBy.Derate:	F_TxtLimitBy := "Derate";
	E_UnitLimitBy.Scaled:	F_TxtLimitBy := "유닛별 값 축소";
	E_UnitLimitBy.BatDir:	F_TxtLimitBy := "배터리 방향";
	E_UnitLimitBy.BatLimit:	F_TxtLimitBy := "배터리 한도";
	E_UnitLimitBy.SLimit:	F_TxtLimitBy := "피상전력";
	E_UnitLimitBy.ModeSwitch:	F_TxtLimitBy := "모드 전환 중";
	E_UnitLimitBy.WaitManualCmd:	F_TxtLimitBy := "새 Manual 지령 대기";
	E_UnitLimitBy.UnitRule:	F_TxtLimitBy := "유닛 제한 모듈";
ELSE
	F_TxtLimitBy := "?";
END_CASE

END_FUNCTION

// ---- 10_Core/70_Diag/F_TxtSeq.TcPOU
FUNCTION F_TxtSeq : WSTRING(31)		// 유닛 시퀀스 문구
VAR_INPUT
	i_e		: E_UnitSeq;
END_VAR

CASE i_e OF
	E_UnitSeq.Unknown:	F_TxtSeq := "알 수 없음";
	E_UnitSeq.Stopped:	F_TxtSeq := "정지";
	E_UnitSeq.WaitBat:	F_TxtSeq := "배터리 투입 대기";
	E_UnitSeq.Standby:	F_TxtSeq := "Standby";
	E_UnitSeq.WaitPermit:	F_TxtSeq := "기동 조건 대기";
	E_UnitSeq.ToRun:	F_TxtSeq := "Run 명령 중";
	E_UnitSeq.Running:	F_TxtSeq := "운전";
	E_UnitSeq.StopRamp:	F_TxtSeq := "정지 램프";
	E_UnitSeq.ToStop:	F_TxtSeq := "정지 명령 중";
ELSE
	F_TxtSeq := "?";
END_CASE

END_FUNCTION

// ---- 10_Core/70_Diag/F_TxtOpMode.TcPOU
FUNCTION F_TxtOpMode : WSTRING(31)		// 운전 모드 문구
VAR_INPUT
	i_e		: E_OpMode;
END_VAR

CASE i_e OF
	E_OpMode.Auto:	F_TxtOpMode := "Auto";
	E_OpMode.Manual:	F_TxtOpMode := "Manual";
ELSE
	F_TxtOpMode := "?";
END_CASE

END_FUNCTION

// ---- 10_Core/70_Diag/FB_AliveRecorder.TcPOU
FUNCTION_BLOCK FB_AliveRecorder		// 마지막 동작 시각을 1 s마다 갱신 (파일 저장은 FB_PersistSave) → 시작할 때 "직전 동작, 꺼져 있던 시간"을 FB_EventLog에 알림 (UPS 신호 없음. 기록은 FB_EventLog가 함)
VAR_IN_OUT
	iq_nLastAlive	: ULINT;			// PERSISTENT: 마지막 동작 시각 (FILETIME 모양, 현지 시각, 100 ns). 글자(iq_sLastAlive)와 같은 출처 FB_LocalSystemTime
	iq_sLastAlive	: STRING(31);		// PERSISTENT: 같은 시각을 현지 시각 글자로
END_VAR
VAR_OUTPUT
	q_bStartLogged	: BOOL;			// 시작 처리를 마침 (이후 1 s마다 시각 갱신)
	q_bStartEvent	: BOOL;			// PMS 시작 (1스캔): FB_EventLog가 기록
	q_sLastAlive	: WSTRING(63);	// 직전 동작 시각 (글자)
	q_sOffTime		: WSTRING(63);	// 꺼져 있던 시간 (글자)
END_VAR
VAR
	_fbLocal		: FB_LocalSystemTime;
	_tonUpdate		: TON;
	_nOffSec		: ULINT;
	_stNowFt		: T_FILETIME;	// 지금 현지 시각 (FILETIME 변환)
	_nNow			: ULINT;			// 지금 현지 시각 (100 ns). 시작 계산·갱신 모두 이 값 하나만 씀
	(* 결함 4 (2026-11-03): 전에는 F_GetSystemTime()(UTC)으로 갱신·비교했는데, 재기동 첫 유효 스캔에서 직전 동작과 1 s 안의 값이 나와
	   꺼져 있던 시간이 0분으로 기록됨 (글자 시각은 맞았음). 글자와 같은 FB_LocalSystemTime 한 곳에서 시각을 얻도록 바꿈 *)
END_VAR

_fbLocal(bEnable := TRUE, dwCycle := 1);
q_bStartEvent := FALSE;
IF _fbLocal.bValid THEN
	_stNowFt := SYSTEMTIME_TO_FILETIME(_fbLocal.systemTime);
	MEMCPY(destAddr := ADR(_nNow), srcAddr := ADR(_stNowFt), n := SIZEOF(_nNow));
END_IF

// 1) 시작 알림: 현지 시각을 처음 얻었을 때 한 번
IF NOT q_bStartLogged AND _fbLocal.bValid THEN
	IF iq_nLastAlive = 0 THEN
		q_sLastAlive := "기록 없음";
		q_sOffTime := "-";
	ELSIF _nNow < iq_nLastAlive THEN
		// 지금이 직전 동작보다 앞 (시각을 뒤로 맞춤 등): 빼면 넘치므로 시간을 내지 않음
		q_sLastAlive	:= STRING_TO_WSTRING(iq_sLastAlive);
		q_sOffTime	:= "알 수 없음 (지금 시각이 직전 동작보다 앞섬)";
	ELSE
		_nOffSec	:= (_nNow - iq_nLastAlive) / 10000000;
		q_sLastAlive	:= STRING_TO_WSTRING(iq_sLastAlive);
		q_sOffTime	:= WCONCAT(TO_WSTRING(_nOffSec / 3600), WCONCAT("시간 ", WCONCAT(TO_WSTRING((_nOffSec MOD 3600) / 60), "분")));
	END_IF
	q_bStartEvent := TRUE;
	q_bStartLogged := TRUE;
END_IF

// 2) 동작 중: 1 s마다 시각 갱신 (메모리만. 파일 저장은 FB_PersistSave가 주기마다)
_tonUpdate(IN := q_bStartLogged AND NOT _tonUpdate.Q, PT := T#1S);
IF _tonUpdate.Q AND _fbLocal.bValid THEN
	iq_nLastAlive := _nNow;
	iq_sLastAlive := SYSTEMTIME_TO_STRING(_fbLocal.systemTime);
END_IF

END_FUNCTION_BLOCK

// ---- 10_Core/02_Util/FB_PersistSave.TcPOU
FUNCTION_BLOCK FB_PersistSave		// PERSISTENT 값을 파일에 저장: 설정이 바뀌면 잠시 뒤 바로, 그리고 주기마다 (PERSISTENT는 정상 종료 때만 저장되므로 직접 씀)
// GVL_PERSIST에 코어 운영 설정을 추가하면 여기 입출력·사본·A_CopyShadow·비교에도 추가한다 (안 넣으면 주기 저장만 됨)
// 현장 모듈 설정 묶음(g_stModuleSet)은 주소·크기로 받아 통째로 비교 → 현장에서 모듈 설정을 늘려도 여기는 안 고침
VAR_INPUT
	i_tPeriod		: TIME := T#60S;	// 주기 저장 (재기동 기록 시각처럼 계속 바뀌는 값)
	i_tSettle		: TIME := T#1S;		// 설정이 바뀐 뒤 이 시간 동안 더 안 바뀌면 저장 (연속 입력을 한 번에)
	i_bSaveNow		: BOOL;				// 바로 저장 요청 (상승 에지)
	i_pModuleSet	: PVOID;			// 현장 모듈 설정 묶음 주소 (ADR(GVL_PERSIST.g_stModuleSet)). 0 = 없음
	i_nModuleSetSize	: UDINT;		// 그 크기 (SIZEOF). GVL_PARAM.MODULE_SET_BYTES보다 크면 비교 안 함 (주기 저장만)
END_VAR
VAR_IN_OUT
	(* 바뀌면 바로 저장할 운영 설정 (GVL_PERSIST). 값은 바꾸지 않음 (VAR_IN_OUT: 저장할 메모리 주소를 비교에 씀) *)
	iq_aeOpMode		: ARRAY[1..GVL_PARAM.UNIT_COUNT] OF E_OpMode;
	iq_astGroupSet	: ARRAY[1..GVL_PARAM.GROUP_COUNT] OF ST_GroupSet;
	iq_astManualPolicy: ARRAY[1..GVL_PARAM.GROUP_COUNT] OF ST_ManualPolicy;
	iq_astSourceReg	: ARRAY[1..GVL_PARAM.SOURCE_COUNT] OF ST_SourceReg;
	iq_astLimitReg	: ARRAY[1..GVL_PARAM.LIMIT_COUNT] OF ST_ModuleReg;
	iq_astPermitReg	: ARRAY[1..GVL_PARAM.PERMIT_COUNT] OF ST_ModuleReg;
	iq_astCompReg	: ARRAY[1..GVL_PARAM.COMP_COUNT] OF ST_ModuleReg;
	iq_astRuleCfg	: ARRAY[1..GVL_PARAM.RULE_COUNT] OF ST_RuleCfg;
	iq_astOutputCfg	: ARRAY[1..GVL_PARAM.OUTPUT_COUNT] OF ST_OutputCfg;
	iq_astUnitRuleReg	: ARRAY[1..GVL_PARAM.UNIT_RULE_COUNT] OF ST_RuleTargetReg;
	iq_astBatRuleReg	: ARRAY[1..GVL_PARAM.BAT_RULE_COUNT] OF ST_RuleTargetReg;
	iq_stCmdFilter	: ST_CmdFilterSet;
	iq_stManualCmdSet	: ST_ManualCmdSet;
	iq_stSeqSet		: ST_SeqSet;
	iq_stBrokerWatch	: ST_BrokerWatchSet;	// [9번 수정 2026-11-09: 추가]
END_VAR
VAR_OUTPUT
	q_bBusy			: BOOL;
	q_bError		: BOOL;				// 마지막 저장 실패
	q_nErrorId		: UDINT;
	q_nSaveCount	: UDINT;			// 성공한 저장 횟수 (PLC 시작 후)
	q_bChangeWait	: BOOL;				// 설정이 바뀌어 저장 대기 중
	q_bModuleSetTooBig	: BOOL;			// 모듈 설정 묶음이 MODULE_SET_BYTES보다 큼: 바뀌어도 바로 저장 안 됨 (GVL_PARAM.MODULE_SET_BYTES를 늘림)
	q_bSetChanged	: BOOL;				// 바뀐 운영 설정을 저장하기 시작함 (1스캔, 기록용)
	q_sSetChanged	: WSTRING(63);		// 그때 바뀐 설정 이름 (마지막 저장 뒤 바뀐 것 모두, 길면 잘림)
END_VAR
VAR
	_fbWrite		: FB_WritePersistentData;
	_tonPeriod		: TON;
	_tonSettle		: TON;
	_rtSaveNow		: R_TRIG;
	_ftBusy			: F_TRIG;
	_bInit			: BOOL;
	_bPending		: BOOL;				// 저장해야 함 (진행 중인 저장이 끝나면 시작)
	_bStart			: BOOL;				// 저장 시작 (한 스캔)
	(* 지난 스캔 사본: 바뀜 확인용 *)
	_aeOpMode		: ARRAY[1..GVL_PARAM.UNIT_COUNT] OF E_OpMode;
	_astGroupSet	: ARRAY[1..GVL_PARAM.GROUP_COUNT] OF ST_GroupSet;
	_astManualPolicy: ARRAY[1..GVL_PARAM.GROUP_COUNT] OF ST_ManualPolicy;
	_astSourceReg	: ARRAY[1..GVL_PARAM.SOURCE_COUNT] OF ST_SourceReg;
	_astLimitReg	: ARRAY[1..GVL_PARAM.LIMIT_COUNT] OF ST_ModuleReg;
	_astPermitReg	: ARRAY[1..GVL_PARAM.PERMIT_COUNT] OF ST_ModuleReg;
	_astCompReg		: ARRAY[1..GVL_PARAM.COMP_COUNT] OF ST_ModuleReg;
	_astRuleCfg		: ARRAY[1..GVL_PARAM.RULE_COUNT] OF ST_RuleCfg;
	_astOutputCfg	: ARRAY[1..GVL_PARAM.OUTPUT_COUNT] OF ST_OutputCfg;
	_astUnitRuleReg	: ARRAY[1..GVL_PARAM.UNIT_RULE_COUNT] OF ST_RuleTargetReg;
	_astBatRuleReg	: ARRAY[1..GVL_PARAM.BAT_RULE_COUNT] OF ST_RuleTargetReg;
	_stCmdFilter	: ST_CmdFilterSet;
	_stManualCmdSet	: ST_ManualCmdSet;
	_stSeqSet		: ST_SeqSet;
	_stBrokerWatch	: ST_BrokerWatchSet;
	_abModuleSet	: ARRAY[0..GVL_PARAM.MODULE_SET_BYTES - 1] OF BYTE;	// 모듈 설정 묶음 사본
	_dwChanged		: DWORD;			// 마지막 저장 뒤 바뀐 설정 (비트 = M_ChangedText 순서)
END_VAR
VAR_TEMP
	bChanged		: BOOL;
	dwNow			: DWORD;			// 이번 스캔에 바뀐 설정
END_VAR

// 모듈 설정 묶음 크기 (첫 스캔 사본 복사보다 먼저: 크면 복사하지 않음)
q_bModuleSetTooBig := i_nModuleSetSize > GVL_PARAM.MODULE_SET_BYTES;

// 첫 스캔: 불러온 값을 기준으로 삼음 (저장 안 함)
IF NOT _bInit THEN
	A_CopyShadow();
	_bInit := TRUE;
END_IF

// 1) 운영 설정이 바뀌었는지 (사본과 메모리 비교)
dwNow := 0;
IF MEMCMP(ADR(iq_aeOpMode), ADR(_aeOpMode), SIZEOF(_aeOpMode)) <> 0 THEN dwNow := dwNow OR 16#00001; END_IF
IF MEMCMP(ADR(iq_astGroupSet), ADR(_astGroupSet), SIZEOF(_astGroupSet)) <> 0 THEN dwNow := dwNow OR 16#00002; END_IF
IF MEMCMP(ADR(iq_astManualPolicy), ADR(_astManualPolicy), SIZEOF(_astManualPolicy)) <> 0 THEN dwNow := dwNow OR 16#00004; END_IF
IF MEMCMP(ADR(iq_astSourceReg), ADR(_astSourceReg), SIZEOF(_astSourceReg)) <> 0 THEN dwNow := dwNow OR 16#00008; END_IF
IF MEMCMP(ADR(iq_astLimitReg), ADR(_astLimitReg), SIZEOF(_astLimitReg)) <> 0 THEN dwNow := dwNow OR 16#00010; END_IF
IF MEMCMP(ADR(iq_astPermitReg), ADR(_astPermitReg), SIZEOF(_astPermitReg)) <> 0 THEN dwNow := dwNow OR 16#00020; END_IF
IF MEMCMP(ADR(iq_astCompReg), ADR(_astCompReg), SIZEOF(_astCompReg)) <> 0 THEN dwNow := dwNow OR 16#00040; END_IF
IF MEMCMP(ADR(iq_astRuleCfg), ADR(_astRuleCfg), SIZEOF(_astRuleCfg)) <> 0 THEN dwNow := dwNow OR 16#00100; END_IF
IF MEMCMP(ADR(iq_astOutputCfg), ADR(_astOutputCfg), SIZEOF(_astOutputCfg)) <> 0 THEN dwNow := dwNow OR 16#00200; END_IF
IF MEMCMP(ADR(iq_astUnitRuleReg), ADR(_astUnitRuleReg), SIZEOF(_astUnitRuleReg)) <> 0 THEN dwNow := dwNow OR 16#00400; END_IF
IF MEMCMP(ADR(iq_astBatRuleReg), ADR(_astBatRuleReg), SIZEOF(_astBatRuleReg)) <> 0 THEN dwNow := dwNow OR 16#00800; END_IF
IF MEMCMP(ADR(iq_stCmdFilter), ADR(_stCmdFilter), SIZEOF(_stCmdFilter)) <> 0 THEN dwNow := dwNow OR 16#02000; END_IF
IF MEMCMP(ADR(iq_stManualCmdSet), ADR(_stManualCmdSet), SIZEOF(_stManualCmdSet)) <> 0 THEN dwNow := dwNow OR 16#04000; END_IF
IF MEMCMP(ADR(iq_stSeqSet), ADR(_stSeqSet), SIZEOF(_stSeqSet)) <> 0 THEN dwNow := dwNow OR 16#08000; END_IF
IF MEMCMP(ADR(iq_stBrokerWatch), ADR(_stBrokerWatch), SIZEOF(_stBrokerWatch)) <> 0 THEN dwNow := dwNow OR 16#20000; END_IF
IF i_pModuleSet <> 0 AND i_nModuleSetSize > 0 AND NOT q_bModuleSetTooBig THEN
	IF MEMCMP(i_pModuleSet, ADR(_abModuleSet), i_nModuleSetSize) <> 0 THEN dwNow := dwNow OR 16#10000; END_IF
END_IF
bChanged := dwNow <> 0;
_dwChanged := _dwChanged OR dwNow;
IF bChanged THEN
	A_CopyShadow();
	q_bChangeWait := TRUE;
	_tonSettle(IN := FALSE);		// 또 바뀌면 대기 시간을 다시 셈
END_IF
_tonSettle(IN := q_bChangeWait, PT := i_tSettle);

// 2) 저장할 때: 바뀐 뒤 잠잠해짐 / 요청 / 주기
_rtSaveNow(CLK := i_bSaveNow);
_tonPeriod(IN := NOT _tonPeriod.Q, PT := i_tPeriod);
q_bSetChanged := FALSE;
IF _tonSettle.Q OR _rtSaveNow.Q OR _tonPeriod.Q THEN
	_bPending		:= TRUE;
	q_bChangeWait	:= FALSE;
	IF _dwChanged <> 0 THEN		// 바뀐 설정을 저장함 → 기록 (FB_EventLog)
		q_bSetChanged	:= TRUE;
		q_sSetChanged	:= M_ChangedText(_dwChanged);
		_dwChanged		:= 0;
	END_IF
END_IF

// 3) 저장 (진행 중이면 끝난 뒤 한 번 더)
_bStart := _bPending AND NOT _fbWrite.BUSY AND NOT _bStart;
IF _bStart THEN
	_bPending := FALSE;
END_IF
_fbWrite(NETID := '', PORT := TwinCAT_SystemInfoVarList._AppInfo.AdsPort, START := _bStart, TMOUT := T#5S);
_ftBusy(CLK := _fbWrite.BUSY);
IF _ftBusy.Q THEN
	q_bError	:= _fbWrite.ERR;
	q_nErrorId	:= _fbWrite.ERRID;
	IF NOT _fbWrite.ERR THEN
		q_nSaveCount := q_nSaveCount + 1;
	END_IF
END_IF
q_bBusy := _fbWrite.BUSY;

METHOD PRIVATE M_ChangedText : WSTRING(63)	// 바뀐 설정 비트 → 이름 (쉼표로 이음, 길면 잘림)
VAR_INPUT
	i_dwMask	: DWORD;
END_VAR
VAR
	i	: INT;
	sName	: WSTRING(31);
	sAll	: WSTRING(255);
END_VAR
sAll := "";
FOR i := 0 TO 17 DO
	IF (SHR(i_dwMask, i) AND 16#1) <> 0 THEN
		CASE i OF
			0:	sName := "운전 모드";
			1:	sName := "그룹 설정";
			2:	sName := "Manual 정책";
			3:	sName := "지령원 등록";
			4:	sName := "제한 등록";
			5:	sName := "기동 조건 등록";
			6:	sName := "보정 등록";
			8:	sName := "보호 규칙";
			9:	sName := "출력 규칙";
			10:	sName := "유닛 제한 등록";
			11:	sName := "버스 제한 등록";
			13:	sName := "명령 필터";
			14:	sName := "Manual 지령 거르기";
			15:	sName := "시퀀스";
			16:	sName := "모듈 설정";
			17:	sName := "브로커 감시";
		ELSE
			sName := "?";
		END_CASE
		IF sAll <> "" THEN
			sAll := WCONCAT(sAll, ", ");
		END_IF
		sAll := WCONCAT(sAll, sName);
	END_IF
END_FOR
M_ChangedText := sAll;
END_METHOD

ACTION A_CopyShadow:
// 지난 스캔 사본 갱신
_aeOpMode		:= iq_aeOpMode;
_astGroupSet	:= iq_astGroupSet;
_astManualPolicy	:= iq_astManualPolicy;
_astSourceReg	:= iq_astSourceReg;
_astLimitReg	:= iq_astLimitReg;
_astPermitReg	:= iq_astPermitReg;
_astCompReg		:= iq_astCompReg;
_astRuleCfg		:= iq_astRuleCfg;
_astOutputCfg	:= iq_astOutputCfg;
_astUnitRuleReg	:= iq_astUnitRuleReg;
_astBatRuleReg	:= iq_astBatRuleReg;
_stCmdFilter	:= iq_stCmdFilter;
_stManualCmdSet	:= iq_stManualCmdSet;
_stSeqSet		:= iq_stSeqSet;
_stBrokerWatch	:= iq_stBrokerWatch;
IF i_pModuleSet <> 0 AND i_nModuleSetSize > 0 AND NOT q_bModuleSetTooBig THEN
	MEMCPY(ADR(_abModuleSet), i_pModuleSet, i_nModuleSetSize);
END_IF
END_ACTION

END_FUNCTION_BLOCK

// ---- 10_Core/70_Diag/FB_ConfigCheck.TcPOU
FUNCTION_BLOCK FB_ConfigCheck		// 매 스캔 고정 설정(GVL_SITE 구성·모듈 ID)을 점검. 운전 중 바꾸는 설정은 FB_SettingGuard가 되돌리고, 되돌릴 정상값이 없을 때만 여기서 오류. 오류가 있으면 q_bConfigOk = FALSE → 장비 쓰기 전부 차단. 오류 문구(앞 10건)를 내고, 기록은 FB_EventLog
VAR_IN_OUT CONSTANT
	iq_astUnitCfg	: ARRAY[1..GVL_PARAM.UNIT_COUNT] OF ST_UnitCfg;
	iq_astBmsCfg	: ARRAY[1..GVL_PARAM.BMS_COUNT] OF ST_BmsCfg;
	iq_astGroupCfg	: ARRAY[1..GVL_PARAM.GROUP_COUNT] OF ST_GroupCfg;
	iq_astPointCfg	: ARRAY[1..GVL_PARAM.POINT_COUNT] OF ST_PointCfg;
END_VAR
VAR_IN_OUT CONSTANT
	iq_abUnitInstalled	: ARRAY[1..GVL_PARAM.UNIT_COUNT] OF BOOL;	// FB_ModuleList: 미설치 유닛은 정격 점검에서 뺌
END_VAR
VAR_INPUT
	i_bModuleSetTooBig	: BOOL;		// 현장 모듈 설정 묶음이 GVL_PARAM.MODULE_SET_BYTES보다 큼 (바로 저장·되돌리기 안 됨)
	i_bSetNoGood	: BOOL;			// 운전 중 바꾸는 설정 값이 잘못됐는데 되돌릴 정상값이 없음 (FB_SettingGuard.q_bNoGood)
	i_sSetNoGood	: WSTRING(63);	// 그 설정과 이유
	i_stRedSet		: ST_RedSet;	// 이중화 설정 (GVL_SITE.RED_SET)
	i_eRedRole		: E_RedRole;	// 이 PLC의 역할 (GVL_IF.g_eRedRole)
END_VAR
VAR_IN_OUT
	iq_aipModule	: ARRAY[1..GVL_PARAM.MODULE_MAX] OF I_Module;	// 등록된 모듈 전부 (FB_ModuleList): 모듈 ID 겹침·0 점검
	iq_aipCtrlMode	: ARRAY[1..GVL_PARAM.CTRL_MODE_COUNT] OF I_ControlMode;	// 제어 모드 (GVL_SITE.g_aipCtrlMode1). 모듈 목록에 없어 따로 점검 [2번 수정 2026-11-09: 추가]
END_VAR
VAR_OUTPUT
	q_bConfigOk		: BOOL;			// 설정 오류 없음. FALSE면 디스패처·보조 출력·시퀀서 명령을 막음
	q_nErrors		: UINT;			// 이번 스캔 오류 수
	q_asErrors		: ARRAY[1..10] OF WSTRING(63);	// 이번 스캔 오류 문구 (앞 10건, 나머지 칸은 빈 문구)
END_VAR
VAR
	_nErrCount		: UINT;								// 이번 스캔 오류 수
	_tonRedReading	: TON;								// 이중화 역할을 못 정한 시간 (Reading, 명세 RED-03 v2.56)
END_VAR
VAR_TEMP
	i				: UINT;
	k				: UINT;
	n				: UINT;
	bZeroId			: BOOL;			// 등록된 모듈 중 ID 0이 있음
	anModuleId			: ARRAY[1..GVL_PARAM.MODULE_MAX] OF UINT;		// 등록된 모듈 ID (0 = 빈 칸)
	anModeId			: ARRAY[1..GVL_PARAM.CTRL_MODE_COUNT] OF UINT;	// 제어 모드 ID (0 = 빈 칸)
END_VAR

_nErrCount := 0;
FOR k := 1 TO 10 DO
	q_asErrors[k] := "";
END_FOR


FOR i := 1 TO GVL_PARAM.UNIT_COUNT DO
	IF iq_astUnitCfg[i].nPcs < 1 OR iq_astUnitCfg[i].nPcs > GVL_PARAM.PCS_COUNT THEN M_AddConfigError(F_TxtNum("UNIT_CFG nPcs 범위 밖: 유닛 ", i)); END_IF
	IF iq_astUnitCfg[i].nSub < 1 OR iq_astUnitCfg[i].nSub > GVL_PARAM.MAX_SUB THEN M_AddConfigError(F_TxtNum("UNIT_CFG nSub 범위 밖: 유닛 ", i)); END_IF
	IF iq_astUnitCfg[i].nBatGroup > GVL_PARAM.BAT_COUNT THEN M_AddConfigError(F_TxtNum("UNIT_CFG nBatGroup 범위 밖: 유닛 ", i)); END_IF
	IF iq_astUnitCfg[i].nGroup < 1 OR iq_astUnitCfg[i].nGroup > GVL_PARAM.GROUP_COUNT THEN M_AddConfigError(F_TxtNum("UNIT_CFG nGroup 범위 밖: 유닛 ", i)); END_IF
	IF iq_abUnitInstalled[i] AND iq_astUnitCfg[i].fPRated <= 0 THEN		// 미설치 유닛(PCS 칸 빈 것)은 정격을 안 봄
		 M_AddConfigError(F_TxtNum("UNIT_CFG fPRated 0 이하: 유닛 ", i)); END_IF
	FOR k := i + 1 TO GVL_PARAM.UNIT_COUNT DO
		IF iq_astUnitCfg[i].nPcs = iq_astUnitCfg[k].nPcs AND iq_astUnitCfg[i].nSub = iq_astUnitCfg[k].nSub THEN
			M_AddConfigError(F_TxtNum("UNIT_CFG 같은 PCS·nSub 중복: 유닛 ", k));
		END_IF
	END_FOR
END_FOR
FOR i := 1 TO GVL_PARAM.BMS_COUNT DO
	IF iq_astBmsCfg[i].nBatGroup < 1 OR iq_astBmsCfg[i].nBatGroup > GVL_PARAM.BAT_COUNT THEN M_AddConfigError(F_TxtNum("BMS_CFG nBatGroup 범위 밖: BMS ", i)); END_IF
END_FOR
FOR i := 1 TO GVL_PARAM.GROUP_COUNT DO
	IF iq_astGroupCfg[i].nPccPoint > GVL_PARAM.POINT_COUNT THEN M_AddConfigError(F_TxtNum("GROUP_CFG nPccPoint 범위 밖: 그룹 ", i)); END_IF
END_FOR
FOR i := 1 TO GVL_PARAM.POINT_COUNT DO
	FOR k := 1 TO GVL_PARAM.POINT_TERM_MAX DO
		IF iq_astPointCfg[i].astTerm[k].nMeter > GVL_PARAM.METER_COUNT THEN M_AddConfigError(F_TxtNum("POINT_CFG nMeter 범위 밖: 계측점 ", i)); END_IF
	END_FOR
END_FOR
// 모듈 ID 겹침·0: 등록된 모듈 목록(FB_ModuleList)으로 비교
n := GVL_PARAM.MODULE_MAX;
bZeroId := FALSE;
FOR i := 1 TO n DO
	anModuleId[i] := 0;
	IF iq_aipModule[i] <> 0 THEN
		anModuleId[i] := iq_aipModule[i].ModuleId;
		bZeroId := bZeroId OR anModuleId[i] = 0;
	END_IF
END_FOR
// 모듈 ID 0은 코어 예약 번호 (등록된 칸인데 0이면 오류)
IF bZeroId THEN
	M_AddConfigError("모듈 ID 0 (코어 예약 번호)인 등록 있음");
END_IF
FOR i := 1 TO n DO
	FOR k := i + 1 TO n DO
		IF anModuleId[i] <> 0 AND anModuleId[i] = anModuleId[k] THEN
			M_AddConfigError(F_TxtNum("모듈 ID 겹침: ", anModuleId[i]));
		END_IF
	END_FOR
END_FOR
// [2번 수정 2026-11-09: 추가] 제어 모드 ID: 0 (코어 예약), 제어 모드끼리 겹침, 등록 모듈과 겹침. 제어 모드는 지령원(관리자) 안의 부품이라 FB_ModuleList에 없어 원래 점검하지 않았음
FOR i := 1 TO GVL_PARAM.CTRL_MODE_COUNT DO
	anModeId[i] := 0;
	IF iq_aipCtrlMode[i] <> 0 THEN
		anModeId[i] := iq_aipCtrlMode[i].ModuleId;
		IF anModeId[i] = 0 THEN
			M_AddConfigError(F_TxtNum("제어 모드 ID 0 (코어 예약 번호): 칸 ", i));
		END_IF
	END_IF
END_FOR
FOR i := 1 TO GVL_PARAM.CTRL_MODE_COUNT DO
	IF anModeId[i] <> 0 THEN
		FOR k := i + 1 TO GVL_PARAM.CTRL_MODE_COUNT DO
			IF anModeId[i] = anModeId[k] THEN
				M_AddConfigError(F_TxtNum("제어 모드 ID 겹침: ", anModeId[i]));
			END_IF
		END_FOR
		FOR k := 1 TO n DO
			IF anModeId[i] = anModuleId[k] THEN
				M_AddConfigError(F_TxtNum("제어 모드 ID가 등록 모듈과 겹침: ", anModeId[i]));
			END_IF
		END_FOR
	END_IF
END_FOR

(* 운전 중 바꾸는 설정 값: 잘못된 값은 FB_SettingGuard가 마지막 정상값으로 되돌림. 되돌릴 정상값이 없을 때(시작부터 잘못)만 설정 오류 *)
IF i_bSetNoGood THEN M_AddConfigError(WCONCAT("설정 값: ", i_sSetNoGood)); END_IF
IF i_bModuleSetTooBig THEN M_AddConfigError("모듈 설정 묶음이 MODULE_SET_BYTES보다 큼"); END_IF
// 이중화: Net ID 두 개가 있어야 하고 서로 달라야 함, 이 PLC Net ID가 둘 중 하나여야 함
IF i_stRedSet.bUse THEN
	IF i_stRedSet.sPrimaryNetId = '' OR i_stRedSet.sSecondaryNetId = '' OR i_stRedSet.sPrimaryNetId = i_stRedSet.sSecondaryNetId THEN
		M_AddConfigError("RED_SET: Primary·Secondary Net ID를 서로 다르게 적어야 함");
	ELSIF i_eRedRole = E_RedRole.NoMatch THEN
		M_AddConfigError("RED_SET: 이 PLC Net ID가 Primary·Secondary와 다름");
	END_IF
END_IF
// 이중화 역할을 10초 넘게 못 정함: Net ID 읽기 실패(PRG_Redundancy.fbGetNetId) 또는 RedundancyTask 정지. PlcTask에서 봐서 그 태스크가 멈춰도 알 수 있음 (명세 RED-03 v2.56)
_tonRedReading(IN := i_stRedSet.bUse AND i_eRedRole = E_RedRole.Reading, PT := T#10S);
IF _tonRedReading.Q THEN M_AddConfigError("RED_SET: 10초 넘게 역할을 못 정함 (Net ID 읽기·RedundancyTask)"); END_IF

q_nErrors	:= _nErrCount;
q_bConfigOk	:= _nErrCount = 0;

METHOD PRIVATE M_AddConfigError
VAR_INPUT
	i_sText		: WSTRING(63);
END_VAR
// 오류 하나를 모음 (기록은 FB_EventLog가 내용이 바뀔 때만)
_nErrCount := _nErrCount + 1;
IF _nErrCount <= 10 THEN
	q_asErrors[_nErrCount] := i_sText;
END_IF
END_METHOD

END_FUNCTION_BLOCK

// ---- 10_Core/70_Diag/FB_SettingGuard.TcPOU
FUNCTION_BLOCK FB_SettingGuard	// 운전 중 바꾸는 설정 값 지키기: 잘못된 값은 받지 않고 마지막 정상값으로 되돌림 (GVL_PERSIST에 다시 씀 → 화면·저장값도 정상값)
// 대상: 코어 설정(명령 필터·Manual 지령 거르기·시퀀스), 등록·출력·규칙 설정(번호 범위, 묶음 통째로), 현장 모듈 설정 묶음(각 모듈 M_CheckSet)
// 처음부터(PMS 시작 때) 잘못이면 되돌릴 정상값이 없으므로 q_bNoGood → FB_ConfigCheck가 설정 오류로 올림 (고치면 그 값이 정상값이 됨)
// 모듈 설정은 묶음 통째로 되돌림 (같은 때 바꾼 다른 모듈 값도 되돌아감). 되돌린 스캔은 q_bRestored → MAIN이 모듈에 다시 넘김
// MAIN ⓪에서 모듈 설정 넘기기·모듈 목록 다음, FB_ConfigCheck 앞에 부름
VAR_INPUT
	i_pModuleSet	: PVOID;		// 현장 모듈 설정 묶음 주소 (ADR(GVL_PERSIST.g_stModuleSet))
	i_nModuleSetSize	: UDINT;	// 그 크기. GVL_PARAM.MODULE_SET_BYTES보다 크면 모듈 설정은 되돌리지 않음 (설정 오류는 FB_ConfigCheck)
END_VAR
VAR_IN_OUT
	iq_stCmdFilter	: ST_CmdFilterSet;		// GVL_PERSIST.g_stCmdFilter (잘못이면 되돌려 씀)
	iq_stManualCmdSet	: ST_ManualCmdSet;	// GVL_PERSIST.g_stManualCmdSet
	iq_stSeqSet		: ST_SeqSet;			// GVL_PERSIST.g_stSeqSet
	iq_astGroupSet	: ARRAY[1..GVL_PARAM.GROUP_COUNT] OF ST_GroupSet;	// GVL_PERSIST.g_astGroupSet (램프율이 숫자가 아니면 되돌림). [결함 13 수정 2026-11-04: 추가]
	iq_aipModule	: ARRAY[1..GVL_PARAM.MODULE_MAX] OF I_Module;	// 등록된 모듈 (FB_ModuleList)
	(* 등록·출력·규칙 설정 (GVL_PERSIST, 운전 중 HMI로 바꿈): 번호가 범위 밖이면 묶음 통째로 되돌림 *)
	iq_astOutputCfg	: ARRAY[1..GVL_PARAM.OUTPUT_COUNT] OF ST_OutputCfg;
	iq_astRuleCfg	: ARRAY[1..GVL_PARAM.RULE_COUNT] OF ST_RuleCfg;
	iq_astSourceReg	: ARRAY[1..GVL_PARAM.SOURCE_COUNT] OF ST_SourceReg;
	iq_astLimitReg	: ARRAY[1..GVL_PARAM.LIMIT_COUNT] OF ST_ModuleReg;
	iq_astPermitReg	: ARRAY[1..GVL_PARAM.PERMIT_COUNT] OF ST_ModuleReg;
	iq_astCompReg	: ARRAY[1..GVL_PARAM.COMP_COUNT] OF ST_ModuleReg;
	iq_astUnitRuleReg	: ARRAY[1..GVL_PARAM.UNIT_RULE_COUNT] OF ST_RuleTargetReg;
	iq_astBatRuleReg	: ARRAY[1..GVL_PARAM.BAT_RULE_COUNT] OF ST_RuleTargetReg;
	(* 위 점검에 쓰는 등록 배열 (모듈이 등록된 칸만 봄) *)
	iq_aipLimit		: ARRAY[1..GVL_PARAM.LIMIT_COUNT] OF I_LimitRule;
	iq_aipPermit	: ARRAY[1..GVL_PARAM.PERMIT_COUNT] OF I_StartPermit;
	iq_aipComp		: ARRAY[1..GVL_PARAM.COMP_COUNT] OF I_Compensator;
	iq_aipRule		: ARRAY[1..GVL_PARAM.RULE_COUNT] OF I_ProtectionRule;
END_VAR
VAR_OUTPUT
	q_bRejected		: BOOL;			// 이번 스캔에 잘못된 값을 되돌림 (1스캔, 기록용)
	q_sRejected		: WSTRING(63);	// 되돌린 설정과 이유 (마지막)
	q_bRestored		: BOOL;			// 이번 스캔에 모듈 설정 묶음을 되돌림 → MAIN이 모듈에 다시 넘김
	q_bNoGood		: BOOL;			// 잘못된 값인데 되돌릴 정상값이 없음 (시작부터 잘못) → 설정 오류
	q_sNoGood		: WSTRING(63);	// 그 설정과 이유
	q_bModuleSetTooBig	: BOOL;		// 모듈 설정 묶음이 GVL_PARAM.MODULE_SET_BYTES보다 큼 (되돌리기·바로 저장 안 됨) → FB_ConfigCheck가 설정 오류로 올림
END_VAR
VAR
	_stCmdFilter	: ST_CmdFilterSet;		// 마지막 정상값
	_stManualCmdSet	: ST_ManualCmdSet;
	_stSeqSet		: ST_SeqSet;
	_abModuleSet	: ARRAY[0..GVL_PARAM.MODULE_SET_BYTES - 1] OF BYTE;
	_bGoodCmdFilter	: BOOL;			// 정상값을 가진 적 있음
	_bGoodManualCmdSet	: BOOL;
	_bGoodSeqSet	: BOOL;
	_astGroupSet	: ARRAY[1..GVL_PARAM.GROUP_COUNT] OF ST_GroupSet;	// 마지막 정상값 [결함 13 수정 2026-11-04: 추가]
	_bGoodGroupSet	: BOOL;
	_bGoodModuleSet	: BOOL;
	(* 등록·출력·규칙 설정 마지막 정상값 *)
	_astOutputCfg	: ARRAY[1..GVL_PARAM.OUTPUT_COUNT] OF ST_OutputCfg;
	_astRuleCfg		: ARRAY[1..GVL_PARAM.RULE_COUNT] OF ST_RuleCfg;
	_astSourceReg	: ARRAY[1..GVL_PARAM.SOURCE_COUNT] OF ST_SourceReg;
	_astLimitReg	: ARRAY[1..GVL_PARAM.LIMIT_COUNT] OF ST_ModuleReg;
	_astPermitReg	: ARRAY[1..GVL_PARAM.PERMIT_COUNT] OF ST_ModuleReg;
	_astCompReg		: ARRAY[1..GVL_PARAM.COMP_COUNT] OF ST_ModuleReg;
	_astUnitRuleReg	: ARRAY[1..GVL_PARAM.UNIT_RULE_COUNT] OF ST_RuleTargetReg;
	_astBatRuleReg	: ARRAY[1..GVL_PARAM.BAT_RULE_COUNT] OF ST_RuleTargetReg;
	_bGoodReg		: BOOL;
	(* A_CheckReg가 씀 (액션은 VAR에 둔 값만 씀) *)
	_sRegErr		: WSTRING(63);	// 등록·출력·규칙 설정 오류 문구 (빈 문구 = 정상, 처음 걸린 것 하나)
	_nRegIdx		: UINT;
	_nRegMax		: UINT;			// 보호 규칙 대상 번호 상한 (범위마다)
END_VAR
VAR_TEMP
	i		: UINT;
	sErr	: WSTRING(63);
	bModuleSetOk	: BOOL;		// 묶음 크기가 되돌릴 수 있는 크기
END_VAR

q_bRejected	:= FALSE;
q_bRestored	:= FALSE;
q_bNoGood	:= FALSE;
q_sNoGood	:= "";

(* 코어 설정 *)
sErr := M_CheckCmdFilter(iq_stCmdFilter);
IF sErr = "" THEN
	_stCmdFilter := iq_stCmdFilter;	_bGoodCmdFilter := TRUE;
ELSIF _bGoodCmdFilter THEN
	iq_stCmdFilter := _stCmdFilter;	M_Reject(WCONCAT("명령 필터: ", sErr));
ELSE
	M_NoGood(WCONCAT("g_stCmdFilter ", sErr));
END_IF

sErr := M_CheckManualCmdSet(iq_stManualCmdSet);
IF sErr = "" THEN
	_stManualCmdSet := iq_stManualCmdSet;	_bGoodManualCmdSet := TRUE;
ELSIF _bGoodManualCmdSet THEN
	iq_stManualCmdSet := _stManualCmdSet;	M_Reject(WCONCAT("Manual 지령 거르기: ", sErr));
ELSE
	M_NoGood(WCONCAT("g_stManualCmdSet ", sErr));
END_IF

sErr := M_CheckSeqSet(iq_stSeqSet);
IF sErr = "" THEN
	_stSeqSet := iq_stSeqSet;	_bGoodSeqSet := TRUE;
ELSIF _bGoodSeqSet THEN
	iq_stSeqSet := _stSeqSet;	M_Reject(WCONCAT("시퀀스: ", sErr));
ELSE
	M_NoGood(WCONCAT("g_stSeqSet ", sErr));
END_IF

(* 그룹 설정: 램프율 REAL이 숫자인지 ([결함 13 수정 2026-11-04: 추가. 범위는 FB_ShapePath가 씀)] *)
sErr := "";
FOR i := 1 TO GVL_PARAM.GROUP_COUNT DO
	IF sErr = "" AND NOT (F_RealOk(iq_astGroupSet[i].fRampUp) AND F_RealOk(iq_astGroupSet[i].fRampDn) AND F_RealOk(iq_astGroupSet[i].fRampResume)) THEN
		sErr := F_TxtNum("램프율 숫자 아님: 그룹 ", i);
	END_IF
END_FOR
IF sErr = "" THEN
	_astGroupSet := iq_astGroupSet;	_bGoodGroupSet := TRUE;
ELSIF _bGoodGroupSet THEN
	iq_astGroupSet := _astGroupSet;	M_Reject(WCONCAT("그룹 설정: ", sErr));
ELSE
	FOR i := 1 TO GVL_PARAM.GROUP_COUNT DO	// 되돌릴 값이 없으면 숫자 아닌 칸만 0 (램프 없음)으로
		IF NOT F_RealOk(iq_astGroupSet[i].fRampUp) THEN iq_astGroupSet[i].fRampUp := 0; END_IF
		IF NOT F_RealOk(iq_astGroupSet[i].fRampDn) THEN iq_astGroupSet[i].fRampDn := 0; END_IF
		IF NOT F_RealOk(iq_astGroupSet[i].fRampResume) THEN iq_astGroupSet[i].fRampResume := 0; END_IF
	END_FOR
	M_NoGood(WCONCAT("g_astGroupSet ", sErr));
END_IF

(* 등록·출력·규칙 설정: 번호 범위 (틀리면 묶음 통째로 되돌림) *)
A_CheckReg();
sErr := _sRegErr;
IF sErr = "" THEN
	A_SaveReg();	_bGoodReg := TRUE;
ELSIF _bGoodReg THEN
	A_RestoreReg();	M_Reject(sErr);
ELSE
	M_NoGood(sErr);
END_IF

(* 모듈 설정: 모듈이 스스로 점검 (MAIN이 이 스캔에 넘긴 값). 처음 걸린 모듈 문구 *)
sErr := "";
FOR i := 1 TO GVL_PARAM.MODULE_MAX DO
	IF sErr = "" AND iq_aipModule[i] <> 0 THEN
		sErr := iq_aipModule[i].M_CheckSet();
		IF sErr <> "" THEN
			sErr := WCONCAT(WCONCAT(STRING_TO_WSTRING(iq_aipModule[i].ModuleName), ": "), sErr);
		END_IF
	END_IF
END_FOR
q_bModuleSetTooBig := i_nModuleSetSize > GVL_PARAM.MODULE_SET_BYTES;
bModuleSetOk := i_pModuleSet <> 0 AND i_nModuleSetSize > 0 AND NOT q_bModuleSetTooBig;
IF sErr = "" THEN
	IF bModuleSetOk THEN
		MEMCPY(ADR(_abModuleSet), i_pModuleSet, i_nModuleSetSize);
		_bGoodModuleSet := TRUE;
	END_IF
ELSIF bModuleSetOk AND _bGoodModuleSet THEN
	MEMCPY(i_pModuleSet, ADR(_abModuleSet), i_nModuleSetSize);
	q_bRestored := TRUE;
	M_Reject(sErr);
ELSE
	M_NoGood(sErr);
END_IF

METHOD PRIVATE M_Reject	// 잘못된 값을 되돌림 (기록용 출력)
VAR_INPUT
	i_sText	: WSTRING(63);
END_VAR
q_bRejected	:= TRUE;
q_sRejected	:= i_sText;
END_METHOD

METHOD PRIVATE M_NoGood	// 잘못됐는데 되돌릴 정상값이 없음 → 설정 오류
VAR_INPUT
	i_sText	: WSTRING(63);
END_VAR
IF NOT q_bNoGood THEN
	q_sNoGood := i_sText;		// 처음 것 하나
END_IF
q_bNoGood := TRUE;
END_METHOD

METHOD PRIVATE M_CheckCmdFilter : WSTRING(63)	// 빈 문구 = 정상
VAR_INPUT
	i_stSet	: ST_CmdFilterSet;
END_VAR
M_CheckCmdFilter := "";
IF NOT F_RealOk(i_stSet.fBadFactor) THEN	// [결함 13 수정 2026-11-04: 숫자 아님(NaN·무한대)은 비교 전에 거름]
	M_CheckCmdFilter := "fBadFactor 숫자 아님";
ELSIF i_stSet.bBadValue AND i_stSet.fBadFactor <= 1.0 THEN
	M_CheckCmdFilter := "fBadFactor 1 이하";
END_IF
END_METHOD

METHOD PRIVATE M_CheckManualCmdSet : WSTRING(63)	// 빈 문구 = 정상
VAR_INPUT
	i_stSet	: ST_ManualCmdSet;
END_VAR
M_CheckManualCmdSet := "";
IF NOT F_RealOk(i_stSet.fDirBand) THEN	// [결함 13 수정 2026-11-04]
	M_CheckManualCmdSet := "fDirBand 숫자 아님";
ELSIF i_stSet.fDirBand < 0.0 OR i_stSet.fDirBand > 100.0 THEN
	M_CheckManualCmdSet := "fDirBand 범위 밖 (0~100 %)";
END_IF
END_METHOD

METHOD PRIVATE M_CheckSeqSet : WSTRING(63)	// 빈 문구 = 정상
VAR_INPUT
	i_stSet	: ST_SeqSet;
END_VAR
M_CheckSeqSet := "";
IF i_stSet.tWritePeriod = T#0S THEN
	M_CheckSeqSet := "tWritePeriod 0";
ELSIF i_stSet.stPcs.tCmdConfirm = T#0S OR i_stSet.stPcs.tStopRetry = T#0S THEN
	M_CheckSeqSet := "PCS 확인 시간 0 (tCmdConfirm·tStopRetry)";
ELSIF NOT F_RealOk(i_stSet.stPcs.fStopDonePct) THEN	// [결함 13 수정 2026-11-04]
	M_CheckSeqSet := "fStopDonePct 숫자 아님";
ELSIF i_stSet.stPcs.fStopDonePct < 0.0 OR i_stSet.stPcs.fStopDonePct > 100.0 THEN
	M_CheckSeqSet := "fStopDonePct 범위 밖 (0~100 %)";
ELSIF i_stSet.stPcs.bStopRamp AND i_stSet.stPcs.tStopRampMax = T#0S THEN
	M_CheckSeqSet := "tStopRampMax 0 (정지 램프 켬)";
ELSIF i_stSet.stBat.tConfirm = T#0S OR i_stSet.stBat.tOpenRetry = T#0S THEN
	M_CheckSeqSet := "배터리 확인 시간 0 (tConfirm·tOpenRetry)";
END_IF
END_METHOD

ACTION A_CheckReg:
// 등록·출력·규칙 설정의 번호 범위 → _sRegErr (빈 문구 = 정상, 처음 걸린 것 하나)
_sRegErr := "";
// [결함 13 수정 2026-11-04: 규칙·출력 칸 REAL(fThreshold, stProt.fPPct·fQPct)이 숫자인지 먼저 (아래 범위 비교·규칙 판단에서 NaN이면 FPU 예외)]
FOR _nRegIdx := 1 TO GVL_PARAM.RULE_COUNT DO
	IF _sRegErr = "" AND NOT (F_RealOk(iq_astRuleCfg[_nRegIdx].fThreshold) AND F_RealOk(iq_astRuleCfg[_nRegIdx].stProt.fPPct) AND F_RealOk(iq_astRuleCfg[_nRegIdx].stProt.fQPct)) THEN
		_sRegErr := F_TxtNum("g_astRuleCfg 값 숫자 아님: 규칙 ", _nRegIdx);
	END_IF
END_FOR
FOR _nRegIdx := 1 TO GVL_PARAM.OUTPUT_COUNT DO
	IF _sRegErr = "" AND NOT F_RealOk(iq_astOutputCfg[_nRegIdx].fThreshold) THEN _sRegErr := F_TxtNum("g_astOutputCfg fThreshold 숫자 아님: 출력 ", _nRegIdx); END_IF
END_FOR
// 보조 출력 칸: 장비·점 번호
FOR _nRegIdx := 1 TO GVL_PARAM.OUTPUT_COUNT DO
	IF _sRegErr = "" AND iq_astOutputCfg[_nRegIdx].nAux > GVL_PARAM.AUX_COUNT THEN _sRegErr := F_TxtNum("g_astOutputCfg nAux 범위 밖: 출력 ", _nRegIdx); END_IF
	IF _sRegErr = "" AND iq_astOutputCfg[_nRegIdx].nAux > 0 AND (iq_astOutputCfg[_nRegIdx].nPoint < 1 OR iq_astOutputCfg[_nRegIdx].nPoint > GVL_PARAM.AUX_DO_MAX) THEN
		_sRegErr := F_TxtNum("g_astOutputCfg nPoint 범위 밖: 출력 ", _nRegIdx);
	END_IF
END_FOR
// 보호 규칙 대상: 범위에 맞는 번호인지 (0 = 범위 안 전부. 틀리면 보호가 걸려도 조치 대상이 없음)
FOR _nRegIdx := 1 TO GVL_PARAM.RULE_COUNT DO
	IF _sRegErr = "" AND iq_aipRule[_nRegIdx] <> 0 AND_THEN (iq_astRuleCfg[_nRegIdx].stProt.bAuto OR iq_astRuleCfg[_nRegIdx].stProt.bManual) THEN
		CASE iq_astRuleCfg[_nRegIdx].eScope OF
			E_ProtScope.Unit:		_nRegMax := GVL_PARAM.UNIT_COUNT;
			E_ProtScope.Bms:		_nRegMax := GVL_PARAM.BMS_COUNT;
			E_ProtScope.BatGroup:	_nRegMax := GVL_PARAM.BAT_COUNT;
			E_ProtScope.Group:		_nRegMax := GVL_PARAM.GROUP_COUNT;
		ELSE
			_nRegMax := 0;				// Site: 대상 번호 안 씀
		END_CASE
		IF _nRegMax > 0 AND iq_astRuleCfg[_nRegIdx].nTarget > _nRegMax THEN
			_sRegErr := F_TxtNum("g_astRuleCfg nTarget 범위 밖: 규칙 ", _nRegIdx);
		END_IF
		// 표준 대응 조치: 배터리 조치는 PCS 정지·비상정지와만 (시퀀서가 PCS 정지 확인 뒤 배터리를 엶), P·Q 상한은 0~100 %
		IF _sRegErr = "" AND iq_astRuleCfg[_nRegIdx].stProt.eBatAction <> E_BatAction.None
			AND NOT (iq_astRuleCfg[_nRegIdx].stProt.ePcsAction = E_PcsAction.Stop OR iq_astRuleCfg[_nRegIdx].stProt.ePcsAction = E_PcsAction.EStop) THEN
			_sRegErr := F_TxtNum("g_astRuleCfg 배터리 조치는 PCS 정지·비상정지와만: 규칙 ", _nRegIdx);
		END_IF
		IF _sRegErr = "" AND (iq_astRuleCfg[_nRegIdx].stProt.fPPct < 0.0 OR iq_astRuleCfg[_nRegIdx].stProt.fPPct > 100.0
			OR iq_astRuleCfg[_nRegIdx].stProt.fQPct < 0.0 OR iq_astRuleCfg[_nRegIdx].stProt.fQPct > 100.0) THEN
			_sRegErr := F_TxtNum("g_astRuleCfg P·Q 상한 0~100 % 밖: 규칙 ", _nRegIdx);
		END_IF
	END_IF
END_FOR
// 등록의 대상 제어 그룹 (0 = 모든 그룹)
FOR _nRegIdx := 1 TO GVL_PARAM.SOURCE_COUNT DO
	IF _sRegErr = "" AND iq_astSourceReg[_nRegIdx].nGroup > GVL_PARAM.GROUP_COUNT THEN _sRegErr := F_TxtNum("g_astSourceReg nGroup 범위 밖: 칸 ", _nRegIdx); END_IF
END_FOR
FOR _nRegIdx := 1 TO GVL_PARAM.LIMIT_COUNT DO
	IF _sRegErr = "" AND iq_astLimitReg[_nRegIdx].nGroup > GVL_PARAM.GROUP_COUNT THEN _sRegErr := F_TxtNum("g_astLimitReg nGroup 범위 밖: 칸 ", _nRegIdx); END_IF
END_FOR
FOR _nRegIdx := 1 TO GVL_PARAM.PERMIT_COUNT DO
	IF _sRegErr = "" AND iq_astPermitReg[_nRegIdx].nGroup > GVL_PARAM.GROUP_COUNT THEN _sRegErr := F_TxtNum("g_astPermitReg nGroup 범위 밖: 칸 ", _nRegIdx); END_IF
END_FOR
FOR _nRegIdx := 1 TO GVL_PARAM.COMP_COUNT DO
	IF _sRegErr = "" AND iq_astCompReg[_nRegIdx].nGroup > GVL_PARAM.GROUP_COUNT THEN _sRegErr := F_TxtNum("g_astCompReg nGroup 범위 밖: 칸 ", _nRegIdx); END_IF
END_FOR
// 유닛 제한·버스 제한의 대상 번호 (0 = 전체)
FOR _nRegIdx := 1 TO GVL_PARAM.UNIT_RULE_COUNT DO
	IF _sRegErr = "" AND iq_astUnitRuleReg[_nRegIdx].nTarget > GVL_PARAM.UNIT_COUNT THEN _sRegErr := F_TxtNum("g_astUnitRuleReg nTarget 범위 밖: 칸 ", _nRegIdx); END_IF
END_FOR
FOR _nRegIdx := 1 TO GVL_PARAM.BAT_RULE_COUNT DO
	IF _sRegErr = "" AND iq_astBatRuleReg[_nRegIdx].nTarget > GVL_PARAM.BAT_COUNT THEN _sRegErr := F_TxtNum("g_astBatRuleReg nTarget 범위 밖: 칸 ", _nRegIdx); END_IF
END_FOR
// 제어 그룹이 2개 이상이면 제한·보정·기동 조건 모듈은 그룹을 지정해야 함 (nGroup 0이면 한 인스턴스가 그룹마다 평가돼 모듈 안 타이머·상태가 섞임 → 그룹마다 인스턴스를 따로 둠)
IF GVL_PARAM.GROUP_COUNT > 1 THEN
	FOR _nRegIdx := 1 TO GVL_PARAM.LIMIT_COUNT DO
		IF _sRegErr = "" AND iq_aipLimit[_nRegIdx] <> 0 AND_THEN (iq_astLimitReg[_nRegIdx].bEnable AND iq_astLimitReg[_nRegIdx].nGroup = 0) THEN _sRegErr := F_TxtNum("g_astLimitReg nGroup 0 (그룹 지정 필요): 칸 ", _nRegIdx); END_IF
	END_FOR
	FOR _nRegIdx := 1 TO GVL_PARAM.PERMIT_COUNT DO
		IF _sRegErr = "" AND iq_aipPermit[_nRegIdx] <> 0 AND_THEN (iq_astPermitReg[_nRegIdx].bEnable AND iq_astPermitReg[_nRegIdx].nGroup = 0) THEN _sRegErr := F_TxtNum("g_astPermitReg nGroup 0 (그룹 지정 필요): 칸 ", _nRegIdx); END_IF
	END_FOR
	FOR _nRegIdx := 1 TO GVL_PARAM.COMP_COUNT DO
		IF _sRegErr = "" AND iq_aipComp[_nRegIdx] <> 0 AND_THEN (iq_astCompReg[_nRegIdx].bEnable AND iq_astCompReg[_nRegIdx].nGroup = 0) THEN _sRegErr := F_TxtNum("g_astCompReg nGroup 0 (그룹 지정 필요): 칸 ", _nRegIdx); END_IF
	END_FOR
END_IF
END_ACTION

ACTION A_SaveReg:
// 등록·출력·규칙 설정을 마지막 정상값으로 저장
_astOutputCfg		:= iq_astOutputCfg;
_astRuleCfg			:= iq_astRuleCfg;
_astSourceReg		:= iq_astSourceReg;
_astLimitReg		:= iq_astLimitReg;
_astPermitReg		:= iq_astPermitReg;
_astCompReg			:= iq_astCompReg;
_astUnitRuleReg		:= iq_astUnitRuleReg;
_astBatRuleReg		:= iq_astBatRuleReg;
END_ACTION

ACTION A_RestoreReg:
// 등록·출력·규칙 설정을 마지막 정상값으로 되돌림 (GVL_PERSIST에 다시 씀)
iq_astOutputCfg		:= _astOutputCfg;
iq_astRuleCfg		:= _astRuleCfg;
iq_astSourceReg		:= _astSourceReg;
iq_astLimitReg		:= _astLimitReg;
iq_astPermitReg		:= _astPermitReg;
iq_astCompReg		:= _astCompReg;
iq_astUnitRuleReg	:= _astUnitRuleReg;
iq_astBatRuleReg	:= _astBatRuleReg;
END_ACTION

END_FUNCTION_BLOCK

// ---- 10_Core/70_Diag/FB_ModuleList.TcPOU
FUNCTION_BLOCK FB_ModuleList	// 등록된 모듈 전부를 한 목록으로 (모듈 ID 점검·이름·이유 문구 찾기는 이 목록만 봄). 유닛·BMS 설치 여부도 냄 (등록 정보)
// 새 등록 배열을 추가하면 여기와 GVL_PARAM.MODULE_MAX만 고침. 칸 순서는 아래 등록 순서, 빈 칸은 0
// 같은 인스턴스를 여러 배열에 등록하면 목록에는 한 번만 (예: 차단기 모듈 = 보호 규칙 + 출력 규칙 2칸, 드라이버 하나가 I_Meter + I_AuxDevice)
VAR_IN_OUT
	iq_aipPcs	: ARRAY[1..GVL_PARAM.PCS_COUNT] OF I_Pcs;
	iq_aipBms	: ARRAY[1..GVL_PARAM.BMS_COUNT] OF I_Bms;
	iq_aipMeter	: ARRAY[1..GVL_PARAM.METER_COUNT] OF I_Meter;
	iq_aipAux	: ARRAY[1..GVL_PARAM.AUX_COUNT] OF I_AuxDevice;
	iq_aipSource	: ARRAY[1..GVL_PARAM.SOURCE_COUNT] OF I_CommandSource;
	iq_aipLimit	: ARRAY[1..GVL_PARAM.LIMIT_COUNT] OF I_LimitRule;
	iq_aipPermit	: ARRAY[1..GVL_PARAM.PERMIT_COUNT] OF I_StartPermit;
	iq_aipComp	: ARRAY[1..GVL_PARAM.COMP_COUNT] OF I_Compensator;
	iq_aipRule	: ARRAY[1..GVL_PARAM.RULE_COUNT] OF I_ProtectionRule;
	iq_aipResp		: ARRAY[1..GVL_PARAM.RULE_COUNT] OF I_ProtResponse;
	iq_aipOutput	: ARRAY[1..GVL_PARAM.OUTPUT_COUNT] OF I_OutputRule;
	iq_aipUnitRule	: ARRAY[1..GVL_PARAM.UNIT_RULE_COUNT] OF I_UnitLimitRule;
	iq_aipBatRule	: ARRAY[1..GVL_PARAM.BAT_RULE_COUNT] OF I_BatLimitRule;
	iq_aipSelPolicy	: ARRAY[1..GVL_PARAM.GROUP_COUNT] OF I_SelectPolicy;
	iq_aipDistPolicy	: ARRAY[1..GVL_PARAM.GROUP_COUNT] OF I_DistPolicy;
	iq_ipAutoGate	: I_Gate;
	iq_ipManualGate	: I_Gate;
END_VAR
VAR_IN_OUT CONSTANT
	iq_astUnitCfg	: ARRAY[1..GVL_PARAM.UNIT_COUNT] OF ST_UnitCfg;
END_VAR
VAR_OUTPUT
	q_aipModule	: ARRAY[1..GVL_PARAM.MODULE_MAX] OF I_Module;	// 등록된 모듈 (같은 인스턴스는 한 번만, 나머지 칸은 0)
	q_abUnitInstalled	: ARRAY[1..GVL_PARAM.UNIT_COUNT] OF BOOL;	// 유닛의 PCS 칸이 등록됨. FALSE = 미설치 (보호·가용·설정 점검에서 뺌)
	q_abBmsInstalled	: ARRAY[1..GVL_PARAM.BMS_COUNT] OF BOOL;	// BMS 칸이 등록됨
END_VAR
VAR
	_n	: UINT;		// 목록에 넣은 칸 수 (M_Add)
END_VAR
VAR_TEMP
	i	: UINT;
	nPcs	: UINT;
END_VAR

_n := 0;
FOR i := 1 TO GVL_PARAM.PCS_COUNT DO M_Add(iq_aipPcs[i]); END_FOR
FOR i := 1 TO GVL_PARAM.BMS_COUNT DO M_Add(iq_aipBms[i]); END_FOR
FOR i := 1 TO GVL_PARAM.METER_COUNT DO M_Add(iq_aipMeter[i]); END_FOR
FOR i := 1 TO GVL_PARAM.AUX_COUNT DO M_Add(iq_aipAux[i]); END_FOR
FOR i := 1 TO GVL_PARAM.SOURCE_COUNT DO M_Add(iq_aipSource[i]); END_FOR
FOR i := 1 TO GVL_PARAM.LIMIT_COUNT DO M_Add(iq_aipLimit[i]); END_FOR
FOR i := 1 TO GVL_PARAM.PERMIT_COUNT DO M_Add(iq_aipPermit[i]); END_FOR
FOR i := 1 TO GVL_PARAM.COMP_COUNT DO M_Add(iq_aipComp[i]); END_FOR
FOR i := 1 TO GVL_PARAM.RULE_COUNT DO M_Add(iq_aipRule[i]); END_FOR
FOR i := 1 TO GVL_PARAM.RULE_COUNT DO M_Add(iq_aipResp[i]); END_FOR
FOR i := 1 TO GVL_PARAM.OUTPUT_COUNT DO M_Add(iq_aipOutput[i]); END_FOR
FOR i := 1 TO GVL_PARAM.UNIT_RULE_COUNT DO M_Add(iq_aipUnitRule[i]); END_FOR
FOR i := 1 TO GVL_PARAM.BAT_RULE_COUNT DO M_Add(iq_aipBatRule[i]); END_FOR
FOR i := 1 TO GVL_PARAM.GROUP_COUNT DO M_Add(iq_aipSelPolicy[i]); END_FOR
FOR i := 1 TO GVL_PARAM.GROUP_COUNT DO M_Add(iq_aipDistPolicy[i]); END_FOR
M_Add(iq_ipAutoGate);
M_Add(iq_ipManualGate);

(* 설치 여부: 칸이 비어 있으면 미설치 *)
FOR i := 1 TO GVL_PARAM.UNIT_COUNT DO
	nPcs := iq_astUnitCfg[i].nPcs;
	q_abUnitInstalled[i] := nPcs >= 1 AND nPcs <= GVL_PARAM.PCS_COUNT AND_THEN iq_aipPcs[nPcs] <> 0;
END_FOR
FOR i := 1 TO GVL_PARAM.BMS_COUNT DO
	q_abBmsInstalled[i] := iq_aipBms[i] <> 0;
END_FOR

METHOD PRIVATE M_Add		// 다음 칸에 모듈을 넣음. 빈 칸이거나 이미 넣은 인스턴스면 0
VAR_INPUT
	i_ipModule	: I_Module;
END_VAR
VAR
	k		: UINT;
	pNew	: POINTER TO BYTE;		// 인스턴스 주소 (같은 인스턴스인지 비교)
	pOld	: POINTER TO BYTE;
	bDup	: BOOL;
END_VAR
_n := _n + 1;
IF _n > GVL_PARAM.MODULE_MAX THEN
	RETURN;
END_IF
q_aipModule[_n] := 0;
IF i_ipModule = 0 THEN
	RETURN;
END_IF
__QUERYPOINTER(i_ipModule, pNew);
FOR k := 1 TO _n - 1 DO
	IF q_aipModule[k] <> 0 THEN
		__QUERYPOINTER(q_aipModule[k], pOld);
		IF pOld = pNew THEN
			bDup := TRUE;
		END_IF
	END_IF
END_FOR
IF NOT bDup THEN
	q_aipModule[_n] := i_ipModule;
END_IF
END_METHOD

END_FUNCTION_BLOCK

// ---- 10_Core/80_Report/FB_Report.TcPOU
FUNCTION_BLOCK FB_Report		// 보고 자리: 코어 결과 → 상위 인터페이스(토탈 인터페이스) 매핑. 보고 전용, 제어는 이 값을 읽지 않음 (R6)
VAR_IN_OUT CONSTANT
	iq_astUnit		: ARRAY[1..GVL_PARAM.UNIT_COUNT] OF ST_UnitState;
	iq_astBms		: ARRAY[1..GVL_PARAM.BMS_COUNT] OF ST_BatState;
	iq_astView		: ARRAY[1..GVL_PARAM.GROUP_COUNT] OF ST_GroupView;
	iq_astAutoPDiag	: ARRAY[1..GVL_PARAM.GROUP_COUNT] OF ST_OutputDiag;
	iq_aeUnitSeq	: ARRAY[1..GVL_PARAM.UNIT_COUNT] OF E_UnitSeq;
	iq_astWritten	: ARRAY[1..GVL_PARAM.UNIT_COUNT] OF ST_PQ;
END_VAR
(* 출력: 인터페이스 구조체가 정해지면 VAR_IN_OUT으로 받아서 채움 *)

(* TODO: 인터페이스 매핑 (인터페이스 버전 확정 후) *)
;

END_FUNCTION_BLOCK

// ---- 20_Module/Common/FB_LocalClock.TcPOU
FUNCTION_BLOCK FB_LocalClock		// 현지 시각 읽기 (TwinCAT Tc2_Utilities FB_LocalSystemTime). 코어는 ST_LocalTime만 보므로 다른 플랫폼은 이 FB만 바꿈
VAR_INPUT
	i_sNetId	: T_AmsNetID := '';		// '' = 이 PLC
	i_nSyncSec	: DWORD := 5;			// 운영체제 시각을 다시 읽는 주기 (s). 사이는 PLC가 셈
END_VAR
VAR_OUTPUT
	q_stTime	: ST_LocalTime;
END_VAR
VAR
	_fbTime		: FB_LocalSystemTime;
END_VAR

_fbTime(sNetID := i_sNetId, bEnable := TRUE, dwCycle := i_nSyncSec);
q_stTime.bValid		:= _fbTime.bValid;
q_stTime.nYear		:= _fbTime.systemTime.wYear;
q_stTime.nMonth		:= _fbTime.systemTime.wMonth;
q_stTime.nDay		:= _fbTime.systemTime.wDay;
q_stTime.nDayOfWeek	:= _fbTime.systemTime.wDayOfWeek;		// 0 = 일요일
q_stTime.nHour		:= _fbTime.systemTime.wHour;
q_stTime.nMinute	:= _fbTime.systemTime.wMinute;
q_stTime.nSecond	:= _fbTime.systemTime.wSecond;

END_FUNCTION_BLOCK

// ---- 20_Module/Ups/FB_UpsConfigApply.TcPOU
FUNCTION_BLOCK FB_UpsConfigApply // EMS config/ups → UPS Holding 설정 쓰기
(* EMS가 내린 주기적·펄스 방전 설정을 UPS에 쓰고 되읽어 확인한다 (UPS 설정). 2026-11-02.
   기반 없음(신규).
   대상: H50~H61, H7, H10 (v2.51). 온도보상(H62~H64)은 스케일 확인 전이라 쓰지 않는다.
   2026-11-16 (명세 v2.14 CF-UPS-01): 간헐충전 H57~H61 추가. H58·H59는 H57이 1이면 전압(0.1 V), 2이면 SOC를
   같은 레지스터에 쓴다. EMS 4칸(전압 2, SOC 2) 중 기준에 맞는 2칸만 쓴다. 기준은 받은 값 → 보관값 → UPS 현재 H57 순.
   - 값 하나라도 범위 밖이면 그 UPS의 이번 설정 전체를 버린다 (BadConfig).
   - is_available=0인 필드와 현재 값이 같은 필드는 쓰지 않는다.
   - BAT Mode가 0(부동충전)일 때만 쓴다. 다른 운전 중이면 끝날 때까지 기다린다.
   - 쓰기 금지 상태에서 받은 설정은 적용하지 않고 버린다 (Disabled). 나중에 허용돼도 옛 값을 쓰지 않음.
   단위: 전류 A → 0.1A, 시간 분·초, 횟수 Cycle. EMS 쪽 단위는 확인 필요.
   2026-11-25 (명세 v2.51 CF-UPS-01): H7 부동 충전 전압·H10 충전 전류 추가 (칸 12·13, 값 × 10). 주소가 이어지지 않아
   칸 → 주소를 ITEM_ADDR 표로 찾는다. 범위: H7 0 초과 UPS_CFG_MAX_VOLTAGE_V 이하, H10 0 초과 UPS_CFG_MAX_CURRENT_A 이하.
   2026-11-23: M_Load가 VAR_IN_OUT(iq_stDesired)을 직접 읽던 것을 입력으로 넘김 (컴파일 경고 제거, 동작 같음)
   2026-11-05 (명세 CF-UPS-02·03): 받은 설정을 보관값(iq_stDesired, GVL_PERSIST)에 남기고,
   i_tRecheck마다 UPS 값을 되읽어 보관값과 다르면 다시 쓴다 (UPS 재기동·PMS 재시작·통신 복구 후 복구).
   UPS 고장(i_bUpsFault)·e-stop 중에는 쓰지 않는다. 2026-11-17: 쓰기 요청(20)·되읽기(30) 단계에서도 매 스캔 다시 보고,
   고장·e-stop·부동충전 아님·데이터 무효면 10단계로 돌아가 기다린다 (실패로 세지 않음). 쓰기가 i_nMaxFail회 연속 실패하면 q_bMismatch를 켜고
   새 설정을 받을 때까지 복구를 멈춘다. *)
VAR_INPUT
	i_bEnable : BOOL; // 장비 쓰기 허용
	i_nRxCount : UDINT; // config/ups 수신 누계
	i_stConfig : ST_UpsConfig_Rx; // 이 UPS의 수신 설정
	i_stState : ST_UpsState; // 장비 상태
	i_stRaw : ST_UpsRaw; // 되읽기용 원본
	i_ipUps : I_Ups; // 쓰기 대상
	i_tTimeout : TIME := T#10S; // 주소 하나의 쓰기·되읽기 제한 시간
	i_bUpsFault : BOOL; // UPS 고장 있음 (보고 Status b6). 켜져 있으면 쓰지 않음
	i_tRecheck : TIME := T#10S; // 보관값과 UPS 값을 비교하는 주기
	i_nMaxFail : UINT := 3; // 연속 실패 허용 횟수. 넘으면 q_bMismatch
END_VAR
VAR_IN_OUT
	iq_stDesired : ST_UpsDesiredSet; // 맞춰 둘 설정 보관값 (GVL_PERSIST.g_astUpsDesired[n])
END_VAR
VAR_OUTPUT
	q_bBusy : BOOL; // 적용 중
	q_eResult : E_UpsResult; // 마지막 적용 결과
	q_nErrorAddress : UINT; // 실패한 H 주소. 0 = 없음
	q_nAppliedRx : UDINT; // 마지막으로 처리한 수신 누계
	q_nWriteCount : UDINT; // 적용한 주소 수 누계
	q_bDesiredChanged : BOOL; // 이 스캔에 보관값을 바꿈 (PERSISTENT 바로 저장 요청)
	q_bMismatch : BOOL; // 설정 불일치 알람: 연속 i_nMaxFail회 실패. 새 설정을 받으면 풀림
	q_nRecoverCount : UDINT; // 복구로 다시 쓴 주소 수 누계
END_VAR
VAR CONSTANT
	ITEM_COUNT : UINT := 14;
	ITEM_ADDR : ARRAY[0..ITEM_COUNT-1] OF UINT := [50, 51, 52, 53, 54, 55, 56, 57, 58, 59, 60, 61, 7, 10]; // 칸 → H 주소. H50~H61, H7, H10 (명세 v2.51)
END_VAR
VAR
	_nStep : UINT;
	_nItem : UINT;
	_nLastRx : UDINT;
	_bBad : BOOL;
	_awTarget : ARRAY[0..ITEM_COUNT-1] OF WORD; // 쓸 값
	_abUse : ARRAY[0..ITEM_COUNT-1] OF BOOL;
	_tonTimeout : TON;
	_tonRecheck : TON; // 비교 주기
	_bRecover : BOOL; // 지금 진행 중인 쓰기가 복구인지 (수신이 아니라)
	_nFail : UINT; // 연속 실패 횟수
	_nCheck : UINT;
END_VAR

_tonTimeout(IN:=_nStep=20 OR _nStep=30, PT:=i_tTimeout);
_tonRecheck(IN:=_nStep=0 AND NOT _tonRecheck.Q, PT:=i_tRecheck);
q_bDesiredChanged:=FALSE;

CASE _nStep OF
	0: // 새 설정 대기
		q_bBusy:=FALSE;
		IF i_nRxCount<>_nLastRx THEN
			_nLastRx:=i_nRxCount;
			q_nErrorAddress:=0;
			IF NOT i_bEnable OR i_ipUps=0 THEN
				q_eResult:=E_UpsResult.Disabled;
				q_nAppliedRx:=_nLastRx;
			ELSE
				M_Load(i_bSavedMode:=iq_stDesired.bValid AND iq_stDesired.abUse[7], i_wSavedMode:=iq_stDesired.awValue[7]);
				IF _bBad THEN
					q_eResult:=E_UpsResult.BadConfig;
					q_nAppliedRx:=_nLastRx;
				ELSE
					// 받은 설정을 보관값으로 남김 (CF-UPS-02)
					iq_stDesired.abUse:=_abUse;
					iq_stDesired.awValue:=_awTarget;
					iq_stDesired.nRxCount:=_nLastRx;
					iq_stDesired.bValid:=TRUE;
					q_bDesiredChanged:=TRUE;
					q_bMismatch:=FALSE;
					_nFail:=0;
					_bRecover:=FALSE;
					q_bBusy:=TRUE;
					q_eResult:=E_UpsResult.Busy;
					_nItem:=0;
					_nStep:=10;
				END_IF
			END_IF
		ELSIF _tonRecheck.Q AND iq_stDesired.bValid AND i_bEnable AND i_ipUps<>0 AND NOT q_bMismatch AND i_stState.bValid THEN
			// 복구 (CF-UPS-03): 보관값과 UPS 값이 다른 칸이 있으면 다시 쓴다
			_abUse:=iq_stDesired.abUse;
			_awTarget:=iq_stDesired.awValue;
			_bRecover:=FALSE;
			FOR _nCheck:=0 TO ITEM_COUNT-1 DO
				IF _abUse[_nCheck] AND i_stRaw.awParam[ITEM_ADDR[_nCheck]]<>_awTarget[_nCheck] THEN
					_bRecover:=TRUE;
				END_IF
			END_FOR
			IF _bRecover THEN
				q_nErrorAddress:=0;
				q_bBusy:=TRUE;
				q_eResult:=E_UpsResult.Busy;
				_nItem:=0;
				_nStep:=10;
			END_IF
		END_IF

	10: // 부동충전 상태에서만 진행
		IF NOT i_bEnable THEN
			q_eResult:=E_UpsResult.Disabled;
			q_nAppliedRx:=_nLastRx;
			_nStep:=0;
		ELSIF i_stState.bValid AND i_stState.nBatMode=0 AND NOT i_bUpsFault AND NOT i_stState.bEmergencyStop THEN
			WHILE _nItem<ITEM_COUNT DO
				IF _abUse[_nItem] AND i_stRaw.awParam[ITEM_ADDR[_nItem]]<>_awTarget[_nItem] THEN EXIT; END_IF
				_nItem:=_nItem+1;
			END_WHILE
			IF _nItem>=ITEM_COUNT THEN
				q_eResult:=E_UpsResult.Accepted;
				q_nAppliedRx:=_nLastRx;
				_nFail:=0;
				_bRecover:=FALSE;
				_nStep:=0;
			ELSE
				_nStep:=20;
			END_IF
		END_IF

	20: // 쓰기 요청
		IF NOT i_bEnable THEN
			q_eResult:=E_UpsResult.Disabled;
			q_nAppliedRx:=_nLastRx;
			_nStep:=0;
		ELSIF i_bUpsFault OR i_stState.bEmergencyStop OR NOT i_stState.bValid OR i_stState.nBatMode<>0 THEN
			_nStep:=10; // 2026-11-17: 기다리는 동안 고장·e-stop 등이 생김 → 쓰지 않고 10단계에서 기다림
		ELSIF i_ipUps.M_SetParameter(UINT_TO_WORD(ITEM_ADDR[_nItem]),_awTarget[_nItem]) THEN
			_nStep:=30;
		ELSIF _tonTimeout.Q THEN
			_nStep:=900;
		END_IF

	30: // 되읽기 확인
		IF i_bUpsFault OR i_stState.bEmergencyStop THEN
			_nStep:=10; // 2026-11-17: 드라이버가 고장·e-stop으로 쓰기를 뺐을 수 있음 → 실패로 세지 않고 다시 기다림
		ELSIF i_stRaw.awParam[ITEM_ADDR[_nItem]]=_awTarget[_nItem] THEN
			q_nWriteCount:=q_nWriteCount+1;
			IF _bRecover THEN q_nRecoverCount:=q_nRecoverCount+1; END_IF
			_nItem:=_nItem+1;
			_nStep:=10;
		ELSIF _tonTimeout.Q THEN
			_nStep:=900;
		END_IF

	900: // 실패. 남은 주소는 쓰지 않음
		q_eResult:=E_UpsResult.CommUnavailable;
		q_nErrorAddress:=ITEM_ADDR[_nItem];
		q_nAppliedRx:=_nLastRx;
		_nFail:=_nFail+1;
		IF _nFail>=i_nMaxFail THEN q_bMismatch:=TRUE; END_IF // 반복을 멈추고 알람
		_bRecover:=FALSE;
		_nStep:=0;
END_CASE

METHOD PRIVATE M_Load
VAR_INPUT
	i_bSavedMode : BOOL; // 보관값에 간헐충전 기준(H57)이 있음 (iq_stDesired.bValid AND abUse[7])
	i_wSavedMode : WORD; // 그 기준 값 (iq_stDesired.awValue[7])
END_VAR
VAR
	nMode : UDINT; // 간헐충전 기준 0 끔 / 1 전압 / 2 SOC (H57)
	bStartAv : BOOL; // 기준에 맞는 시작 칸을 받음
	bEndAv : BOOL; // 기준에 맞는 종료 칸을 받음
	rStart : REAL;
	rEnd : REAL;
	rScale : REAL; // 레지스터 배율 (전압 10, SOC GVL_PARAM.UPS_CFG_SOC_SCALE)
	rMax : REAL; // 상한 (전압 UPS_CFG_MAX_VOLTAGE_V, SOC 100)
END_VAR
_bBad:=FALSE;
_abUse[0]:=i_stConfig.PeriodicTrickleDischargeSetCurrent.is_available<>0;
IF _abUse[0] THEN
	IF i_stConfig.PeriodicTrickleDischargeSetCurrent.value>0.0 AND i_stConfig.PeriodicTrickleDischargeSetCurrent.value<=GVL_PARAM.UPS_CFG_MAX_CURRENT_A THEN
		_awTarget[0]:=REAL_TO_WORD(i_stConfig.PeriodicTrickleDischargeSetCurrent.value*10.0);
	ELSE _bBad:=TRUE; q_nErrorAddress:=50; END_IF
END_IF
_abUse[1]:=i_stConfig.PeriodicTrickleDischargeSetTime.is_available<>0;
IF _abUse[1] THEN
	IF i_stConfig.PeriodicTrickleDischargeSetTime.value>0 AND i_stConfig.PeriodicTrickleDischargeSetTime.value<=GVL_PARAM.UPS_CFG_MAX_MINUTES THEN
		_awTarget[1]:=UDINT_TO_WORD(i_stConfig.PeriodicTrickleDischargeSetTime.value);
	ELSE _bBad:=TRUE; q_nErrorAddress:=51; END_IF
END_IF
_abUse[2]:=i_stConfig.PulseDischargeSetCurrent.is_available<>0;
IF _abUse[2] THEN
	IF i_stConfig.PulseDischargeSetCurrent.value>0.0 AND i_stConfig.PulseDischargeSetCurrent.value<=GVL_PARAM.UPS_CFG_MAX_CURRENT_A THEN
		_awTarget[2]:=REAL_TO_WORD(i_stConfig.PulseDischargeSetCurrent.value*10.0);
	ELSE _bBad:=TRUE; q_nErrorAddress:=52; END_IF
END_IF
_abUse[3]:=i_stConfig.PulseChargeSetCurrent.is_available<>0;
IF _abUse[3] THEN
	IF i_stConfig.PulseChargeSetCurrent.value>0.0 AND i_stConfig.PulseChargeSetCurrent.value<=GVL_PARAM.UPS_CFG_MAX_CURRENT_A THEN
		_awTarget[3]:=REAL_TO_WORD(i_stConfig.PulseChargeSetCurrent.value*10.0);
	ELSE _bBad:=TRUE; q_nErrorAddress:=53; END_IF
END_IF
_abUse[4]:=i_stConfig.PulseDischargeSetTime.is_available<>0;
IF _abUse[4] THEN
	IF i_stConfig.PulseDischargeSetTime.value>0 AND i_stConfig.PulseDischargeSetTime.value<=GVL_PARAM.UPS_CFG_MAX_SECONDS THEN
		_awTarget[4]:=UDINT_TO_WORD(i_stConfig.PulseDischargeSetTime.value);
	ELSE _bBad:=TRUE; q_nErrorAddress:=54; END_IF
END_IF
_abUse[5]:=i_stConfig.PulseChargeSetTime.is_available<>0;
IF _abUse[5] THEN
	IF i_stConfig.PulseChargeSetTime.value>0 AND i_stConfig.PulseChargeSetTime.value<=GVL_PARAM.UPS_CFG_MAX_SECONDS THEN
		_awTarget[5]:=UDINT_TO_WORD(i_stConfig.PulseChargeSetTime.value);
	ELSE _bBad:=TRUE; q_nErrorAddress:=55; END_IF
END_IF
_abUse[6]:=i_stConfig.PulseChargeDischargeSetCycle.is_available<>0;
IF _abUse[6] THEN
	IF i_stConfig.PulseChargeDischargeSetCycle.value>0 AND i_stConfig.PulseChargeDischargeSetCycle.value<=GVL_PARAM.UPS_CFG_MAX_CYCLES THEN
		_awTarget[6]:=UDINT_TO_WORD(i_stConfig.PulseChargeDischargeSetCycle.value);
	ELSE _bBad:=TRUE; q_nErrorAddress:=56; END_IF
END_IF
// H57~H61 간헐충전 (명세 v2.14 CF-UPS-01). H58·H59는 H57 기준에 따라 전압 또는 SOC
_abUse[7]:=i_stConfig.TrickleChargeSetParameter.is_available<>0;
IF _abUse[7] THEN
	IF i_stConfig.TrickleChargeSetParameter.value<=2 THEN
		nMode:=i_stConfig.TrickleChargeSetParameter.value;
		_awTarget[7]:=UDINT_TO_WORD(nMode);
	ELSE _bBad:=TRUE; q_nErrorAddress:=57; END_IF
ELSIF i_bSavedMode THEN
	nMode:=WORD_TO_UDINT(i_wSavedMode);
ELSE
	nMode:=WORD_TO_UDINT(i_stRaw.awParam[57]);
END_IF
_abUse[8]:=FALSE;
_abUse[9]:=FALSE;
bStartAv:=FALSE;
bEndAv:=FALSE;
IF nMode=1 THEN
	bStartAv:=i_stConfig.TrickleChargeSetStartVoltage.is_available<>0;
	bEndAv:=i_stConfig.TrickleChargeSetEndVoltage.is_available<>0;
	rStart:=i_stConfig.TrickleChargeSetStartVoltage.value;
	rEnd:=i_stConfig.TrickleChargeSetEndVoltage.value;
	rScale:=10.0;
	rMax:=GVL_PARAM.UPS_CFG_MAX_VOLTAGE_V;
ELSIF nMode=2 THEN
	bStartAv:=i_stConfig.TrickleChargeSetStartSoc.is_available<>0;
	bEndAv:=i_stConfig.TrickleChargeSetEndSoc.is_available<>0;
	rStart:=i_stConfig.TrickleChargeSetStartSoc.value;
	rEnd:=i_stConfig.TrickleChargeSetEndSoc.value;
	rScale:=GVL_PARAM.UPS_CFG_SOC_SCALE;
	rMax:=100.0;
END_IF
IF nMode=1 OR nMode=2 THEN
	IF _abUse[7] AND NOT (bStartAv AND bEndAv) THEN
		_bBad:=TRUE; q_nErrorAddress:=58; // 기준을 바꿀 때는 시작·종료를 같이 받아야 함
	ELSE
		IF bStartAv AND bEndAv AND rStart>=rEnd THEN _bBad:=TRUE; q_nErrorAddress:=58; END_IF
		IF bStartAv THEN
			IF rStart>0.0 AND rStart<=rMax THEN _abUse[8]:=TRUE; _awTarget[8]:=REAL_TO_WORD(rStart*rScale);
			ELSE _bBad:=TRUE; q_nErrorAddress:=58; END_IF
		END_IF
		IF bEndAv THEN
			IF rEnd>0.0 AND rEnd<=rMax THEN _abUse[9]:=TRUE; _awTarget[9]:=REAL_TO_WORD(rEnd*rScale);
			ELSE _bBad:=TRUE; q_nErrorAddress:=59; END_IF
		END_IF
	END_IF
END_IF
_abUse[10]:=i_stConfig.TrickleChargeSetStartTime.is_available<>0; // EMS 이름은 StartTime, 맵 H60은 간헐충전 종료시간 (분)
IF _abUse[10] THEN
	IF i_stConfig.TrickleChargeSetStartTime.value>0 AND i_stConfig.TrickleChargeSetStartTime.value<=GVL_PARAM.UPS_CFG_MAX_TRICKLE_MINUTES THEN
		_awTarget[10]:=UDINT_TO_WORD(i_stConfig.TrickleChargeSetStartTime.value);
	ELSE _bBad:=TRUE; q_nErrorAddress:=60; END_IF
END_IF
_abUse[11]:=i_stConfig.TrickleChargeSetReStartDay.is_available<>0;
IF _abUse[11] THEN
	IF i_stConfig.TrickleChargeSetReStartDay.value>0 AND i_stConfig.TrickleChargeSetReStartDay.value<=GVL_PARAM.UPS_CFG_MAX_DAYS THEN
		_awTarget[11]:=UDINT_TO_WORD(i_stConfig.TrickleChargeSetReStartDay.value);
	ELSE _bBad:=TRUE; q_nErrorAddress:=61; END_IF
END_IF
// H7 부동 충전 전압·H10 충전 전류 (명세 v2.51 CF-UPS-01). 값 × 10
_abUse[12]:=i_stConfig.FloatChargeSetVoltage.is_available<>0;
IF _abUse[12] THEN
	IF i_stConfig.FloatChargeSetVoltage.value>0.0 AND i_stConfig.FloatChargeSetVoltage.value<=GVL_PARAM.UPS_CFG_MAX_VOLTAGE_V THEN
		_awTarget[12]:=REAL_TO_WORD(i_stConfig.FloatChargeSetVoltage.value*10.0);
	ELSE _bBad:=TRUE; q_nErrorAddress:=7; END_IF
END_IF
_abUse[13]:=i_stConfig.ChargeSetCurrentLimit.is_available<>0;
IF _abUse[13] THEN
	IF i_stConfig.ChargeSetCurrentLimit.value>0.0 AND i_stConfig.ChargeSetCurrentLimit.value<=GVL_PARAM.UPS_CFG_MAX_CURRENT_A THEN
		_awTarget[13]:=REAL_TO_WORD(i_stConfig.ChargeSetCurrentLimit.value*10.0);
	ELSE _bBad:=TRUE; q_nErrorAddress:=10; END_IF
END_IF
END_METHOD

END_FUNCTION_BLOCK

// ---- 20_Module/Ups/FB_UpsCommand.TcPOU
(* EMS UPS 명령 → 세방 UPS 명령 레지스터(0x55) 요청, 온도보상 켜짐 상태 복구 (⑤출력 / 장치: UPS). 2026-11-05.
   기반 없음(신규).
   변경: 없음
   부호·단위: 해당 없음. 명세: C:\gil\UPS\명세서\UPS_명세서.md WR-UPS-01, CF-UPS-03(켜짐 상태). WR-SQ-01은 v2.38에서 폐기
   - 2026-11-12 인터페이스 100.Command: CommandType은 번호 1~26. 번호 n → 세방 맵 명령 주소 99+n (H100~H125)에 0x55
     1 리셋 2 버저 정지 3·4 정류부 ON·OFF 5·6 인버터 ON·OFF 7·8 BBC ON·OFF 9 인버터로 절체 10 바이패스로 절체
     11 부동충전 12 균등충전 13·14 Auto ON·OFF 15 비상 방전 16 주기적 방전 17 펄스 방전 18 방전 취소
     19·20 간헐충전 시작·취소 21·22 온도보상 시작·취소 23·24 ECO 시작·취소 25·26 PRLT 시작·취소
   - 레코드 하나 = 명령 하나. 버전 2의 Delay 대기는 앞에서 FB_EmsCmdGate가 한다
   - 거부: UPS 통신이상이면 모두. UPS 고장(Status b2)이나 e-stop(b3) 중이면 켜기·시작 명령(START_TYPES). 끄기·취소·리셋은 보냄
   - 쓰기 허용(i_bEnable)이 꺼져 있으면 실행하지 않고 Disabled. 장치 명령 1~26, 보고 모드 101 수동·102 자동을 받음
   - 2026-11-17: 드라이버가 바빠 기다리는 동안에도 매 스캔 다시 본다. 고장·e-stop이 생기면 대기 중인 시작 명령을 취소(BadRequest),
     쓰기 허용이 꺼지면 취소(Disabled). 끄기·취소·리셋은 그대로 보낸다
   - Fault 단계 확인은 EMS가 한다 (명세 v2.4). q_bAck는 늘 FALSE
   - 온도보상: 켜 둬야 하는데(iq_stDesired.bTempCompOn) UPS가 꺼져 있으면 i_tRecheck마다 시작 명령을 다시 보낸다.
     i_nMaxFail회 연속으로 켜지지 않으면 q_bEnableMismatch를 켜고 멈춘다. 21·22를 받으면 풀린다 *)
FUNCTION_BLOCK FB_UpsCommand
VAR_INPUT
	i_stCmd			: ST_IfUpsCmd;			// 받은 명령 (번호가 바뀌면 새 명령)
	i_bEnable		: BOOL;					// 장비 쓰기 허용
	i_stUps			: ST_UpsPublish_V1;		// UPS 보고값 (Status b2 고장, b3 e-stop, UPS_ModeStatus b7 온도보상)
	i_bUpsValid		: BOOL;					// UPS 통신 정상
	i_ipUps			: I_Ups;				// 명령 대상
	i_tRequestTimeout : TIME := T#5S;		// 드라이버가 요청을 받지 못하면 실패로 보는 시간
	i_tRecheck		: TIME := T#10S;		// 온도보상 켜짐 상태 확인 주기
	i_nMaxFail		: UINT := 3;			// 켜짐 상태 복구 연속 실패 허용 횟수
END_VAR
VAR_IN_OUT
	iq_stDesired	: ST_UpsDesiredSet;		// 켜짐 상태 보관값 (GVL_PERSIST.g_astUpsDesired[n])
END_VAR
VAR_OUTPUT
	q_bAck				: BOOL;				// Fault 단계 확인. EMS가 하므로 늘 FALSE (v2.4). v2.38부터 MAIN에서 쓰지 않음 (PMS 안 Fault 유지 없앰)
	q_nOperationMode	: UDINT := 1;		// EMS 보고 운전모드: 0 수동(101), 1 자동(102). 시작 기본값 자동
	q_nLastType			: UDINT;			// 마지막으로 받은 명령 번호
	q_eLastResult		: E_UpsResult;		// 마지막 명령 결과
	q_nRejectCount		: UDINT;			// 상태 때문에 거부한 명령 수
	q_nUnknownCount		: UDINT;			// 1~26·101·102 밖의 번호를 받은 수
	q_bDesiredChanged	: BOOL;				// 이 스캔에 켜짐 상태 보관값을 바꿈 (바로 저장 요청)
	q_bEnableMismatch	: BOOL;				// 온도보상 복구 연속 실패 알람
	q_nRestoreCount		: UDINT;			// 온도보상 복구로 시작 명령을 보낸 횟수
END_VAR
VAR
	_nLastSeq		: UDINT;
	_bInit			: BOOL;
	_nPending		: UDINT;				// 드라이버에 넘길 명령 번호 (0 = 없음)
	_tonRequest		: TON;
	_tonRecheck		: TON;
	_nFail			: UINT;
	_bRestoreSent	: BOOL;					// 지난 확인 때 복구 명령을 보냄
	_bFault			: BOOL;
	_bEStop			: BOOL;
	_eCmd			: E_UpsCommand;
	_nNew			: UDINT;
	_bAccepted		: BOOL;
END_VAR
VAR CONSTANT
	MAX_TYPE		: UDINT := 26;		// 번호 1~26 (H100~H125)
	// 고장·e-stop 중 거부하는 켜기·시작 번호: 3 정류부 ON, 5 인버터 ON, 7 BBC ON, 9 인버터로 절체, 11 부동, 12 균등, 13 Auto ON,
	// 15 비상 방전, 16 주기적 방전, 17 펄스 방전, 19 간헐충전, 21 온도보상, 23 ECO, 25 PRLT (비트 n = 번호 n)
	START_TYPES		: DWORD := 16#02ABBAA8;
END_VAR

q_bAck := FALSE;
q_bDesiredChanged := FALSE;
_bFault := i_stUps.Status.2;	// b2 fault
_bEStop := i_stUps.Status.3;	// b3 e-stop

// 처음 스캔: 재시작 전에 받은 명령 번호를 다시 실행하지 않음
IF NOT _bInit THEN
	_bInit := TRUE;
	_nLastSeq := i_stCmd.nSeq;
END_IF

// 1) 새 명령 (1~26 장치, 101 수동·102 자동 보고 모드)
IF i_stCmd.nSeq <> _nLastSeq THEN
	_nLastSeq := i_stCmd.nSeq;
	q_nLastType := i_stCmd.nType;
	_nNew := i_stCmd.nType;
	IF _nNew = 101 OR _nNew = 102 THEN
		// PMS 보고 모드만 변경한다. 세방 Auto ON/OFF(13/14)나 장치 명령은 보내지 않는다.
		IF i_bEnable THEN
			q_nOperationMode := _nNew - 101;
			q_eLastResult := E_UpsResult.Accepted;
		ELSE
			q_eLastResult := E_UpsResult.Disabled;
		END_IF
	ELSIF _nNew = 0 OR _nNew > MAX_TYPE THEN
		q_nUnknownCount := q_nUnknownCount + 1;
		q_eLastResult := E_UpsResult.BadRequest;
	ELSIF NOT i_bUpsValid THEN
		q_nRejectCount := q_nRejectCount + 1;
		q_eLastResult := E_UpsResult.CommUnavailable;
	ELSIF (_bFault OR _bEStop) AND (START_TYPES AND SHL(DWORD#1, UDINT_TO_INT(_nNew))) <> 0 THEN
		q_nRejectCount := q_nRejectCount + 1;	// 고장·e-stop 중 켜기·시작 거부
		q_eLastResult := E_UpsResult.BadRequest;
	ELSIF NOT i_bEnable OR i_ipUps = 0 THEN
		q_eLastResult := E_UpsResult.Disabled;
	ELSE
		_nPending := _nNew;	// 앞의 요청이 남아 있으면 새 명령으로 바꿈 (마지막 명령이 우선)
		q_eLastResult := E_UpsResult.Busy;
	END_IF
END_IF

// 2) 드라이버에 요청. 받아들이면 켜짐 상태 보관값 갱신
_bAccepted := FALSE;
// 2026-11-17: 기다리는 동안 상태가 바뀌면 대기 명령을 취소 (받을 때만 보던 것을 매 스캔 다시 봄)
IF _nPending <> 0 THEN
	IF (_bFault OR _bEStop) AND (START_TYPES AND SHL(DWORD#1, UDINT_TO_INT(_nPending))) <> 0 THEN
		_nPending := 0;
		q_nRejectCount := q_nRejectCount + 1;	// 고장·e-stop이 생겨 시작 명령 취소
		q_eLastResult := E_UpsResult.BadRequest;
	ELSIF NOT i_bEnable OR i_ipUps = 0 THEN
		_nPending := 0;
		q_eLastResult := E_UpsResult.Disabled;
	END_IF
END_IF
_tonRequest(IN := _nPending <> 0, PT := i_tRequestTimeout);
IF _nPending <> 0 THEN
	CASE _nPending OF	// 번호 n → 맵 주소 99+n (E_UpsCommand 값 = 주소)
		1:	_eCmd := E_UpsCommand.Reset;
		2:	_eCmd := E_UpsCommand.BuzzerStop;
		3:	_eCmd := E_UpsCommand.RectifierOn;
		4:	_eCmd := E_UpsCommand.RectifierOff;
		5:	_eCmd := E_UpsCommand.InverterOn;
		6:	_eCmd := E_UpsCommand.InverterOff;
		7:	_eCmd := E_UpsCommand.BbcOn;
		8:	_eCmd := E_UpsCommand.BbcOff;
		9:	_eCmd := E_UpsCommand.ToInverter;
		10:	_eCmd := E_UpsCommand.ToBypass;
		11:	_eCmd := E_UpsCommand.FloatCharge;
		12:	_eCmd := E_UpsCommand.EqualCharge;
		13:	_eCmd := E_UpsCommand.AutoOn;
		14:	_eCmd := E_UpsCommand.AutoOff;
		15:	_eCmd := E_UpsCommand.EmergencyDischarge;
		16:	_eCmd := E_UpsCommand.PeriodicDischarge;
		17:	_eCmd := E_UpsCommand.PulseDischarge;
		18:	_eCmd := E_UpsCommand.CancelDischarge;
		19:	_eCmd := E_UpsCommand.TrickleOn;
		20:	_eCmd := E_UpsCommand.TrickleOff;
		21:	_eCmd := E_UpsCommand.TemperatureOn;
		22:	_eCmd := E_UpsCommand.TemperatureOff;
		23:	_eCmd := E_UpsCommand.EcoOn;
		24:	_eCmd := E_UpsCommand.EcoOff;
		25:	_eCmd := E_UpsCommand.PrltOn;
		26:	_eCmd := E_UpsCommand.PrltOff;
	END_CASE
	IF i_ipUps.M_RequestCommand(_eCmd) THEN
		_bAccepted := TRUE;
		q_eLastResult := E_UpsResult.Accepted;
		CASE _nPending OF
			19:	iq_stDesired.bTrickleOn := TRUE;	q_bDesiredChanged := TRUE;
			20:	iq_stDesired.bTrickleOn := FALSE;	q_bDesiredChanged := TRUE;
			21:	iq_stDesired.bTempCompOn := TRUE;	q_bDesiredChanged := TRUE;	q_bEnableMismatch := FALSE;	_nFail := 0;	_bRestoreSent := FALSE;
			22:	iq_stDesired.bTempCompOn := FALSE;	q_bDesiredChanged := TRUE;	q_bEnableMismatch := FALSE;	_nFail := 0;	_bRestoreSent := FALSE;
		END_CASE
		_nPending := 0;
		_tonRequest(IN := FALSE);
	ELSIF _tonRequest.Q THEN
		_nPending := 0;	// 드라이버가 받지 못함
		q_eLastResult := E_UpsResult.CommUnavailable;
	END_IF
END_IF

// 3) 온도보상 켜짐 상태 복구 (CF-UPS-03)
_tonRecheck(IN := NOT _tonRecheck.Q, PT := i_tRecheck);
IF _tonRecheck.Q AND _nPending = 0 AND NOT _bAccepted THEN
	IF i_stUps.UPS_ModeStatus.7 OR NOT iq_stDesired.bTempCompOn THEN
		_nFail := 0;					// 켜져 있거나 켤 필요 없음
		_bRestoreSent := FALSE;
	ELSIF i_bUpsValid AND i_bEnable AND i_ipUps <> 0 AND NOT _bFault AND NOT _bEStop AND NOT q_bEnableMismatch THEN
		IF _bRestoreSent THEN
			_nFail := _nFail + 1;		// 지난번에 보냈는데 아직 꺼져 있음
		END_IF
		IF _nFail >= i_nMaxFail THEN
			q_bEnableMismatch := TRUE;	// 반복을 멈추고 알람
		ELSIF i_ipUps.M_RequestCommand(E_UpsCommand.TemperatureOn) THEN
			_bRestoreSent := TRUE;
			q_nRestoreCount := q_nRestoreCount + 1;
		END_IF
	END_IF
END_IF

END_FUNCTION_BLOCK

// ---- 20_Module/Report/FB_RptEsolutionBat.TcPOU
FUNCTION_BLOCK FB_RptEsolutionBat // BMS 시스템 값 → BAT 보고값
VAR_INPUT
	i_stState : ST_EsolutionState; // 장비 상태
	i_stRaw : ST_EsolutionRaw; // 랙·모듈 원본
	i_nDeviceIndex : UDINT; // 배터리 번호 (1부터). 랙·모듈 번호도 모두 1부터 [1부터 2026-11-10]
END_VAR
VAR_OUTPUT
	q_stBat : ST_BatPublish_V1; // BAT 보고값
	q_bValid : BOOL; // 유효한 장비 데이터
	q_astRack : ARRAY[1..GVL_PARAM.RACKS_PER_BMS] OF ST_RackPublish_V1; // RACK 보고값
	q_astModule : ARRAY[1..GVL_PARAM.RACKS_PER_BMS*GVL_PARAM.MODULES_PER_RACK] OF ST_ModulePublish_V1; // MODULE 보고값
END_VAR
VAR
	_stEmpty : ST_BatPublish_V1;
	_stRackEmpty : ST_RackPublish_V1;
	_stModuleEmpty : ST_ModulePublish_V1;
	_nLastSeq : UDINT; // 마지막으로 계산한 표본 번호
	_bLastValid : BOOL;
	_bCalculated : BOOL; // 번호를 한 번은 채웠는가 (통신 없는 BMS도 계산)
	_nRack : UINT;
	_nModule : UINT;
	_nCell : UINT;
	_nIndex : UINT;
	_nAnalog : UINT; // Input 50~89 랙 시작 칸
	_nStatus : UINT; // Input 90~179 랙 시작 칸
	_wOperation : WORD; // 랙 운전 상태
	_wCell : WORD; // 셀 전압 (mV)
	_wCellMax : WORD;
	_wCellMin : WORD;
	_fTemp : REAL;
	_fTempMax : REAL;
	_fTempMin : REAL;
	_pCell : POINTER TO REAL;
	_nOnlineRacks : UDINT; // 릴레이 투입 또는 충·방전 중인 랙 수
	_bInitializing : BOOL;
	_bCharging : BOOL;
	_bDischarging : BOOL;
	_wSysAlarm : WORD; // S+0 System Alarm (마스크 적용)
	_wSysWarn : WORD; // S+2 System Warning Status
	_wSysError : WORD; // S+3 System Error Status
	_wModError : WORD; // S+4 Module Error Status
	_wFire : WORD; // S+7 Fire Alarm
	_wLock1 : WORD; // D+11 System Lock Status 1 (상세 받은 랙만)
	_wLock2 : WORD; // D+12 System Lock Status 2 (상세 받은 랙만)
	_wModule : WORD; // S+8 Module Status
	_wErr1 : WORD; // S+5 Error Code 1
	_wErr2 : WORD; // S+6 Error Code 2 (마스크 적용)
	_wSelf1 : WORD; // D+13 Self Test Status 1 (상세 받은 랙만)
	_wSelf2 : WORD; // D+14 Self Test Status 2 (상세 받은 랙만)
	_bRackWarn : BOOL; // 그 랙 Warning 칸 중 0이 아닌 것이 있음
	_bRackFault : BOOL; // 그 랙 Fault 칸 중 0이 아닌 것이 있음
	_nBatWarn1 : UDINT; // BAT Warning1 = 랙 값 OR
	_nBatWarn2 : UDINT; // BAT Warning2 = 랙 값 OR (명세 RD-BAT-02 v2.48)
	_anBatFault : ARRAY[1..5] OF UDINT; // BAT Fault1~5 = 랙 값 OR (v2.37)
END_VAR
VAR CONSTANT
	// 명세 RD-BAT-01 (v2.48): 배터리 eventMap v2 + Warning2 (공유 드라이브 구글 시트 002.이솔루션, 2026-11-24). 칸 하나에 BMS 워드 2개 (첫 워드 b0~, 둘째 워드 b16~), 각 워드 안에서는 정의된 비트만 이어 붙임.
	// 맵 v1.3·v1.4 Bit_List에서 정의된 비트만 남김 (Reserved는 항상 0)
	SYS_ALARM_MASK : WORD := 16#01FF; // S+0 System Alarm b0~8 → Warning1 b16~24
	SYS_WARN_MASK : WORD := 16#03FF; // S+2 System Warning Status b0~9 → Warning1 b0~9
	SYS_ERROR_MASK : WORD := 16#3FFF; // S+3 System Error Status b0~13 → Fault1 b0~13
	MODULE_ERROR_MASK : WORD := 16#07FF; // S+4 Module Error Status b0~10. (v2.48) b0~8 → Fault1 b16~24, b10 → Fault1 b25, b9 Cell V Imbalance Warning → Warning2 b0
	FIRE_MASK : WORD := 16#8001; // S+7 Fire Alarm b0 연기 센서 → Fault2 b0, b15 화재·연기 감지기 → Fault2 b1
	MODULE_STATUS_MASK : WORD := 16#01FF; // S+8 Module Status b0~8. (v2.48) 에러 b1·3·5·7·8 → Fault2 b16~20, 경고 b0·2·4·6 (UV·OV·OT·UT Warning) → Warning2 b1~4
	LOCK1_MASK : WORD := 16#0FCB; // D+11 System Lock Status 1 b0·1·3·6~11 → Fault3 b0~8
	LOCK2_MASK : WORD := 16#FFF3; // D+12 System Lock Status 2 b0·1·4~15 → Fault3 b16~29
	ERROR_CODE2_MASK : WORD := 16#00FF; // S+6 Error Code 2 b0~7 → Fault4 b16~23 (Error Code 1은 b0~15 모두 → Fault4 b0~15)
	SELF1_MASK : WORD := 16#01FF; // D+13 Self Test Status 1 b0~8 → Fault5 b0~8
	SELF2_MASK : WORD := 16#F7FF; // D+14 Self Test Status 2 b0~10·12~15 (b11 Reserved) → Fault5 b16~30
END_VAR

q_stBat := _stEmpty;
q_stBat.DeviceIndex := i_nDeviceIndex;
q_stBat.TotalRackCount := UINT_TO_UDINT(i_stState.nRackCount);
q_stBat.Status := 1; // b0 통신에러
q_bValid := i_stState.bValid;
IF q_bValid THEN
	q_stBat.Heartbeat := WORD_TO_UDINT(i_stState.nHeartbeat); // 하트비트
	q_stBat.Soc := i_stState.fSocPct; // 충전 상태 (%)
	q_stBat.Soh := i_stState.fSohPct; // 건강 상태 (%)
	q_stBat.DcVoltage := i_stState.fVoltageV; // 전체 전압 (V)
	q_stBat.DcCurrent := i_stState.fCurrentA; // 전체 전류 (A)
	q_stBat.ChargeCurrentLimit := i_stState.fChargeCurrentLimitA; // 충전 허용 전류 (A)
	q_stBat.DischargeCurrentLimit := i_stState.fDischargeCurrentLimitA; // 방전 허용 전류 (A)
	q_stBat.ChargePowerLimit := i_stState.fChargeLimitKw; // 충전 허용 전력 (kW)
	q_stBat.DischargePowerLimit := i_stState.fDischargeLimitKw; // 방전 허용 전력 (kW)
	q_stBat.MaxCellVoltage := i_stState.fMaxCellVoltageMv * 0.001; // 최대 셀 전압 (V)
	q_stBat.MinCellVoltage := i_stState.fMinCellVoltageMv * 0.001; // 최소 셀 전압 (V)
	q_stBat.MaxModuleTemperature := i_stState.fMaxCellTemperatureC; // 맵은 Cell Temperature로 표기
	q_stBat.MinModuleTemperature := i_stState.fMinCellTemperatureC;
	// 위치는 맵 형식 [RRMM]: 0512 = 랙 5, 모듈 12
	q_stBat.MaxCellVoltageLocationFromRack := WORD_TO_UDINT(i_stState.nMaxCellVoltageLocation) / 100;
	q_stBat.MaxCellVoltageLocationFromModule := WORD_TO_UDINT(i_stState.nMaxCellVoltageLocation) MOD 100;
	q_stBat.MinCellVoltageLocationFromRack := WORD_TO_UDINT(i_stState.nMinCellVoltageLocation) / 100;
	q_stBat.MinCellVoltageLocationFromModule := WORD_TO_UDINT(i_stState.nMinCellVoltageLocation) MOD 100;
	q_stBat.MaxModuleTempLocationFromRack := WORD_TO_UDINT(i_stState.nMaxCellTemperatureLocation) / 100;
	q_stBat.MaxModuleTempLocationFromModule := WORD_TO_UDINT(i_stState.nMaxCellTemperatureLocation) MOD 100;
	q_stBat.MinModuleTempLocationFromRack := WORD_TO_UDINT(i_stState.nMinCellTemperatureLocation) / 100;
	q_stBat.MinModuleTempLocationFromModule := WORD_TO_UDINT(i_stState.nMinCellTemperatureLocation) MOD 100;
END_IF

